(* IEC 61131-3 sources: daoli-st-library/DL_Motion (part 20) *)

(* ---- FB_DL_UnwinderDiameterCalc.st ---- *)
(*==============================================================================
 * 组件名称 (Component)  : FB_DL_UnwinderDiameterCalc
 * 所属子库 (Sublibrary) : DL_Motion
 * 当前版本 (Version)    : 1.0.0
 * 兼容性 (Platform)     : CODESYS 3.5 / TwinCAT 3 / 汇川 InoProShop / Machine Expert
 *                         仅依赖纯 IEC 61131-3 标准元素，零厂商方言
 * 功能描述 (Function)   : 放卷卷径实时估算：fDia = sqrt(fDiaInit^2 - 4 x thick x
 *                         SigmaLen / pi)，开方委托 FC_DL_NthRoot(2)；按外部累计
 *                         放膜长度增量递推；低于最小卷径 → bSpoolEnd 预警。
 *                         被开方数 < 0（数据矛盾）→ 冻结并报错，不塞伪值。
 * 溯源 (Origin)         : 道莅 clean-room 防御性实现
 * 本文件内含 (Contains) : TYPE E_DL_UnwdErr / FUNCTION_BLOCK FB_DL_UnwinderDiameterCalc
 * 依赖 (Depends)        : DL_MathData/FC_DL_NthRoot
 * 红线自检 (Redline)    : 无外部全局变量、无硬件地址直引 ｜ 全变量中英双语同行注释
 *                         防除零 + 量程钳位 + 非有限值防御 ｜ 枚举成员全部显式赋值
 *                         开方委托不重实现 ｜ 浮点容差比较 ｜ 输出冻结语义显式
 * 错误码表 (Codes)      : 16#0004_0318 就绪
 *                         16#0004_0319 信息级 膜厚非法(已钳制下限)
 *                         16#0004_031A 故障级 长度增量非法(拒绝递推)
 *                         16#0004_031B 故障级 数据矛盾(根号内负值或非有限，冻结输出)
 *                         16#0004_031C 信息级 接近空卷预警
 * 修订历史 (Revision)   : 2026-11-17  v1.0.0  首版入库 · R27 · 阶段三批 3
 * 验收向量 (Acceptance) : 初始卷径 500 mm，膜厚 50 um，累计放膜 1000 m
 *                         → 卷径 = sqrt(500^2 - 4*0.05*1000/3.14159...) ≈ 499.94 mm
 *============================================================================*)

(*-----------------------------------------------------------------------------
 * 枚举: E_DL_UnwdErr（归属 DL_Motion，与 FB_DL_UnwinderDiameterCalc 同文件）
 *----------------------------------------------------------------------------*)
TYPE E_DL_UnwdErr :
(
    eReady      := 16#0004_0318,   // 就绪 / Ready
    eThickClamp := 16#0004_0319,   // 信息级：膜厚非法已钳制下限 / Info: film thickness clamped
    eLenIncrBad := 16#0004_031A,   // 故障级：长度增量非法（放卷长度不允许回退）/ Fault: illegal length increment
    eDataContrad:= 16#0004_031B,   // 故障级：数据矛盾（根号内负值或非有限，冻结）/ Fault: data contradiction, output frozen
    eSpoolEnd   := 16#0004_031C    // 信息级：接近空卷预警 / Info: spool-end warning
);
END_TYPE

(*==============================================================================
 * 功能块: FB_DL_UnwinderDiameterCalc
 * 调用约定: 每个扫描周期无条件调用一次；fWebLen_m 必须为单调不减的累计放膜长度。
 *============================================================================*)
FUNCTION_BLOCK FB_DL_UnwinderDiameterCalc
VAR_INPUT
    fFilmThick_um : REAL;              // 膜厚 [微米]，有效域 5~500 / Film thickness [um]
    fDiaInit_mm   : REAL;              // 初始卷径 [毫米]，有效域 50~1200 / Initial roll diameter [mm]
    fWebLen_m     : REAL;              // 累计放膜长度 [米]（外部积分输入，单调不减）/ Accumulated web length [m]
    fDiaMin_mm    : REAL;              // 最小卷径 [毫米]（空卷预警门限）/ Minimum roll diameter [mm]
    bReset        : BOOL;              // 换卷复位（重新以初始卷径起算）/ Roll-change reset
END_VAR
VAR_OUTPUT
    fDiaNow_mm    : REAL;              // 当前卷径 [毫米] / Current roll diameter [mm]
    bSpoolEnd     : BOOL;              // 接近空卷预警 / Spool-end warning
    eErr          : E_DL_UnwdErr;      // 错误码 / Error code
END_VAR
VAR
    fLenPrev      : REAL;              // 上拍累计长度快照 [米]（增量基准）/ Previous length snapshot [m]
    fLenUse       : REAL;              // 生效累计长度（增量非法时冻结）[米] / Effective accumulated length [m]
    fThickUse_mm  : REAL;              // 生效膜厚（换算毫米，钳位后）[毫米] / Effective thickness in mm [mm]
    fDiaInitUse   : REAL;              // 生效初始卷径（NaN 兜底）[毫米] / Effective initial diameter [mm]
    fLenIncr      : REAL;              // 本拍长度增量 [米] / Length increment this scan [m]
    fRadicand     : LREAL;             // 被开方数 [平方毫米] / Radicand [mm2]
    fRootVal      : LREAL;             // 委托开方输出 [毫米] / Delegate root output [mm]
    bRootOk       : BOOL;              // 委托开方有效标志 / Delegate root validity flag
    bFrozen       : BOOL;              // 输出冻结标志（数据矛盾置位）/ Output frozen flag
    bInit         : BOOL;              // 首扫初始化标志 / First-scan init flag
END_VAR
VAR CONSTANT
    DL_UNWD_THICK_MIN : REAL := 5.0;      // 膜厚下限 [微米] / Thickness lower bound [um]
    DL_UNWD_THICK_MAX : REAL := 500.0;    // 膜厚上限 [微米] / Thickness upper bound [um]
    DL_UNWD_DIA_MIN   : REAL := 50.0;     // 初始卷径下限 [毫米] / Initial diameter lower bound [mm]
    DL_UNWD_DIA_MAX   : REAL := 1200.0;   // 初始卷径上限 [毫米] / Initial diameter upper bound [mm]
    DL_UNWD_UM2MM     : REAL := 0.001;    // 微米换毫米系数 [毫米每微米] / um-to-mm factor [mm per um]
    DL_UNWD_M2MM      : REAL := 1000.0;   // 米换毫米系数 [毫米每米] / m-to-mm factor [mm per m]
    DL_UNWD_FOUR      : REAL := 4.0;      // 面积递推系数 4（4 x thick x len / pi）/ Area recursion factor
    DL_UNWD_PI        : REAL := 3.14159265358979;   // 圆周率 [无量纲] / Pi [dimensionless]
    DL_UNWD_TOL       : REAL := 1.0E-6;   // 浮点比较容差 / Float comparison tolerance
    DL_UNWD_INF_MAX   : REAL := 1.0E30;   // 非有限值判定幅值上限 / Magnitude bound for finite-value check
    DL_UNWD_ZERO      : REAL := 0.0;      // 零值常量，避免裸字面量 / Zero constant
END_VAR

(*------------------------------------------------------------------------------
 * 段 1｜换卷复位：清快照与冻结标志，卷径回初始值
 *----------------------------------------------------------------------------*)
IF bReset THEN
    fLenPrev := fWebLen_m;                         // 快照重置为当前累计长度 / snapshot reset
    fLenUse := fWebLen_m;                          // 累计长度重置 / length reset
    fDiaNow_mm := fDiaInit_mm;                     // 卷径回初始值 / diameter back to initial
    bFrozen := FALSE;                              // 冻结解除 / freeze released
    bSpoolEnd := FALSE;                            // 预警解除 / warning released
    bInit := TRUE;                                 // 视为首扫完成（跳过旧快照）/ treated as initialized
    eErr := E_DL_UnwdErr.eReady;                   // 回就绪码 / back to ready
    RETURN;
END_IF

(*------------------------------------------------------------------------------
 * 段 2｜首扫初始化：建立长度快照基准
 *----------------------------------------------------------------------------*)
IF NOT bInit THEN
    fLenPrev := fWebLen_m;                         // 首扫快照 / first-scan snapshot
    fLenUse := fWebLen_m;                          // 累计长度基准 / length baseline
    bInit := TRUE;                                 // 首扫完成 / first scan done
END_IF

(*------------------------------------------------------------------------------
 * 段 3｜非有限值闸：任一输入 NaN/溢出 → 冻结输出并报数据矛盾（不塞伪值）
 *----------------------------------------------------------------------------*)
IF (fFilmThick_um <> fFilmThick_um) OR (ABS(fFilmThick_um) > DL_UNWD_INF_MAX)
   OR (fDiaInit_mm <> fDiaInit_mm) OR (ABS(fDiaInit_mm) > DL_UNWD_INF_MAX)
   OR (fWebLen_m <> fWebLen_m) OR (ABS(fWebLen_m) > DL_UNWD_INF_MAX)
   OR (fDiaMin_mm <> fDiaMin_mm) OR (ABS(fDiaMin_mm) > DL_UNWD_INF_MAX) THEN
    bFrozen := TRUE;                               // 输出冻结 / output frozen
    eErr := E_DL_UnwdErr.eDataContrad;             // 故障级：数据矛盾（非有限并入）/ fault: data contradiction
    bSpoolEnd := TRUE;                             // 数据矛盾按安全侧预警 / safe-side warning
    RETURN;
END_IF

(*------------------------------------------------------------------------------
 * 段 4｜膜厚钳位（信息级）与初始卷径兜底
 *----------------------------------------------------------------------------*)
eErr := E_DL_UnwdErr.eReady;                       // 预置就绪 / preset ready
fThickUse_mm := fFilmThick_um * DL_UNWD_UM2MM;     // 膜厚换算毫米 [毫米] / thickness to mm
IF fFilmThick_um < DL_UNWD_THICK_MIN THEN
    fThickUse_mm := DL_UNWD_THICK_MIN * DL_UNWD_UM2MM;   // 膜厚下限钳制 / thickness floored
    eErr := E_DL_UnwdErr.eThickClamp;              // 信息级：膜厚非法已钳制 / info: thickness clamped
ELSIF fFilmThick_um > DL_UNWD_THICK_MAX THEN
    fThickUse_mm := DL_UNWD_THICK_MAX * DL_UNWD_UM2MM;   // 膜厚上限钳制 / thickness capped
    eErr := E_DL_UnwdErr.eThickClamp;              // 信息级：膜厚非法已钳制 / info: thickness clamped
END_IF
fDiaInitUse := fDiaInit_mm;                        // 初始卷径工作副本 / initial diameter working copy
IF (fDiaInitUse < DL_UNWD_DIA_MIN) OR (fDiaInitUse > DL_UNWD_DIA_MAX) THEN
    fDiaInitUse := DL_UNWD_DIA_MIN;                // 初始卷径出域按下限兜底（配置防御）/ initial diameter falls back
END_IF

(*------------------------------------------------------------------------------
 * 段 5｜长度增量合法性闸：放卷长度单调不减（容差内视为零增量）
 *----------------------------------------------------------------------------*)
fLenIncr := fWebLen_m - fLenPrev;                  // 本拍增量 [米] / increment this scan [m]
IF fLenIncr < -DL_UNWD_TOL THEN
    bFrozen := TRUE;                               // 增量为负：拒绝递推，冻结输出 / negative increment: reject, freeze
    eErr := E_DL_UnwdErr.eLenIncrBad;              // 故障级：长度增量非法 / fault: illegal increment
    fLenUse := fLenPrev;                           // 冻结到上拍快照 / frozen at previous snapshot
    RETURN;
END_IF
IF fLenIncr < DL_UNWD_ZERO THEN
    fLenIncr := DL_UNWD_ZERO;                      // 容差内微负增量钳零 / tiny negative clamped to zero
END_IF
fLenUse := fLenPrev + fLenIncr;                    // 生效累计长度 [米] / effective length [m]
fLenPrev := fWebLen_m;                             // 快照推进 / snapshot advanced

(*------------------------------------------------------------------------------
 * 段 6｜卷径递推：被开方数 = 初始卷径^2 - 4 x 膜厚 x 累计长度 / pi
 *       被开方数 < 0（数据矛盾：放膜量超过卷料面积）→ 冻结并报故障级
 *----------------------------------------------------------------------------*)
fRadicand := REAL_TO_LREAL(fDiaInitUse * fDiaInitUse)
           - REAL_TO_LREAL(DL_UNWD_FOUR * fThickUse_mm * fLenUse * DL_UNWD_M2MM) / REAL_TO_LREAL(DL_UNWD_PI);   // 被开方数 [平方毫米]（米换毫米链）/ radicand [mm2]
IF (fRadicand <> fRadicand) OR (ABS(fRadicand) > REAL_TO_LREAL(DL_UNWD_INF_MAX)) THEN
    bFrozen := TRUE;                               // 非有限中间量：冻结 / non-finite intermediate: freeze
    eErr := E_DL_UnwdErr.eDataContrad;             // 故障级：数据矛盾 / fault: data contradiction
    bSpoolEnd := TRUE;                             // 安全侧预警 / safe-side warning
    RETURN;
END_IF
IF fRadicand < LREAL#0.0 THEN
    bFrozen := TRUE;                               // 根号内负值：数据矛盾冻结 / negative radicand: freeze
    eErr := E_DL_UnwdErr.eDataContrad;             // 故障级：根号内负值 / fault: negative radicand
    bSpoolEnd := TRUE;                             // 安全侧预警 / safe-side warning
    RETURN;
END_IF

(*------------------------------------------------------------------------------
 * 段 7｜委托开方（FC_DL_NthRoot(2)）与空卷预警
 *----------------------------------------------------------------------------*)
fRootVal := FC_DL_NthRoot(fValue := fRadicand, nRoot := 2, bValid => bRootOk);   // 开方委托 [毫米] / root via delegate [mm]
IF (NOT bRootOk) OR (fRootVal <> fRootVal) OR (ABS(fRootVal) > REAL_TO_LREAL(DL_UNWD_INF_MAX)) THEN
    bFrozen := TRUE;                               // 委托失败：冻结 / delegate failure: freeze
    eErr := E_DL_UnwdErr.eDataContrad;             // 故障级：数据矛盾（委托失败并入，输出同为冻结）/ fault: contradiction
    RETURN;
END_IF
fDiaNow_mm := LREAL_TO_REAL(fRootVal);             // 当前卷径输出 [毫米] / current diameter output [mm]
IF fDiaNow_mm < DL_UNWD_ZERO THEN
    fDiaNow_mm := DL_UNWD_ZERO;                    // 下限防护 / floor guard
END_IF
bSpoolEnd := fDiaNow_mm <= fDiaMin_mm + DL_UNWD_TOL;   // 空卷预警判据（容差比较）/ spool-end predicate
IF bSpoolEnd THEN
    eErr := E_DL_UnwdErr.eSpoolEnd;                // 信息级：接近空卷 / info: spool-end warning
END_IF
END_FUNCTION_BLOCK

(* ---- FB_DL_VelFfGainIdent.st ---- *)
(*==============================================================================
 * 组件名称 (Component)  : FB_DL_VelFfGainIdent
 * 所属子库 (Sublibrary) : DL_Motion
 * 当前版本 (Version)    : 1.0.0
 * 兼容性 (Platform)     : CODESYS 3.5+ / TwinCAT 3 / 汇川 InoProShop / 施耐德 Machine Expert
 *                         仅依赖 Standard.library（TON / R_TRIG），零厂商私有库，
 *                         零轴状态枚举引用（R277）
 * 功能描述 (Function)   : 速度前馈增益辨识。恒速段窗口（bConstVel 电平：上层
 *                         速度指令平坦段）内对 (vFb, vCmd) 做 最小二乘 过原点
 *                         拟合 K = Σ(vFb·vCmd) / Σ(vFb²)（前馈模型 vCmd ≈ K·vFb
 *                         的残差最优解），同步累计残差标准差与样本数；样本充分
 *                         且拟合优度高（残差/信号比小）→ bIdentDone 单拍输出
 *                         fKvf。与 AxisFrictionFf 分工：本件辨识增益不注入
 *                         前馈（R312 模型不内嵌注入语义）。
 * 来源标签 (Origin)     : 自研线（IEC 61131-3 标准语义的道莅防御性实现，clean-room）
 * 分工声明 (Pairing)    : VelFfGainIdent（辨识，本件）↔ AxisFrictionFf（前馈注入，
 *                         既有件）：本件只产出辨识增益与置信指标，不写前馈通道、
 *                         不驱动轴（R298 属主边界）；辨识结果由调用方决定是否
 *                         下装（R312 口径）。
 * 边界语义 (Boundary)   : ① 过原点拟合分母闸：Σ(vFb²) <= eps（恒速段实际零速
 *                         或样本未采）→ 拟合不执行，K 保持上值；
 *                         ② 速度非有限拒收（NaN 自反 + Inf 差判）；
 *                         ③ 置信闸：残差均方根/均值 |vCmd| > fConfRatio
 *                         → 拟合质量不足，bIdentDone 不置位（辨识不可信
 *                         必须可观测，R28 口径）；
 *                         ④ 组态闸：最小样本/置信比/增益钳位域 → 故障。
 * 输出语义 (Fallback)   : 【R191】bConstVel = FALSE → 停止采样，fKvf 保持
 *                         末次辨识值（增益是资产，不随窗口停而清零）；
 *                         eFault 相 → 冻结 + bError = TRUE。
 * 码位     (Codes)      : 按 R297 范式零 16# 码位硬编码；错误出口 BOOL+ENUM(eCause)，
 *                         码位待主控收口统一派号。
 * 红线自检 (Redline)    : 7 项红线已自检：R1 零全局 ✓｜R2 零物理地址 ✓｜R3 纯 IEC ✓
 *                         R4 除零（Σv² eps 闸）/NaN 拒收/组态闸 ✓
 *                         R5 双语同行注释 ✓｜R6 CASE 带 ELSE 兜底迁 eFault ✓
 *                         R7 TON/R_TRIG 段 0 无条件刷新 ✓
 * 验收向量 (Acceptance) : V1 恒速段 vCmd=vFb=200 → K=1.0（容差 1E-6）；
 *                         V2 vFb 恒为 vCmd 的 0.8 倍 → K=1.25；
 *                         V3 零速恒速段（vFb≈0）→ 分母闸生效，K 保持上值；
 *                         V4 残差比超阈 → bIdentDone 不置位。
 * 修订历史 (Revision)   : 2026-11-20  v1.0.0  R49 首版（批 4 · 序号 17）
 *==============================================================================*)
TYPE E_DL_VfiState :
(
    eIdle  := 0,                             (* 待使能 / Idle *)
    eLearn := 10,                            (* 恒速段采样与拟合 / Learning *)
    eFault := 90                             (* 故障锁存相 / Fault latched phase *)
);
END_TYPE

TYPE E_DL_VfiCause :
(
    eNone       := 0,                        (* 无故障成因 / No cause *)
    eCfgIllegal := 1,                        (* 组态非法：样本/置信比越域 / Illegal config *)
    ePhaseBad   := 2                         (* 非法相位兜底 / Illegal phase fallback *)
);
END_TYPE

FUNCTION_BLOCK FB_DL_VelFfGainIdent
VAR_INPUT
    fVelCmd    : LREAL := 0.0;               (* 速度指令反馈快照 [mm/s] / Velocity command snapshot *)
    fVelFb     : LREAL := 0.0;               (* 实际速度反馈快照 [mm/s] / Velocity feedback snapshot *)
    bConstVel  : BOOL := FALSE;              (* 恒速段电平（上层速度平坦段判据直连）[-] / Constant-velocity window level *)
    nMinSample : INT := 64;                  (* 最小辨识样本数，域 8..100000 [点] / Min identification samples *)
    fConfRatio : LREAL := 0.1;               (* 置信比门限（残差 RMS / 均值|vCmd|），域 (0,1) [-] / Confidence ratio gate *)
    bEnable    : BOOL := TRUE;               (* 辨识使能 [-] / Enable *)
    bReset     : BOOL := FALSE;              (* 复位命令，上升沿清累计与锁存（fKvf 保留）[-] / Reset command *)
END_VAR
VAR_OUTPUT
    fKvf       : LREAL;                      (* 辨识速度前馈增益（末次有效值保持）[-] / Identified velocity ff gain *)
    nSampleCnt : INT;                        (* 本轮累计样本数 [点] / Sample count this round *)
    fResidRms  : LREAL;                      (* 跟随残差均方根（拟合质量）[mm/s] / Residual RMS *)
    bIdentDone : BOOL;                       (* 本轮辨识完成单拍位（质量闸通过才置位）[-] / Round-done single-scan pulse *)
    bIdentFail : BOOL;                       (* 本轮辨识质量不足锁存位（复位沿清）[-] / Round-quality-fail latch *)
    eState     : E_DL_VfiState;              (* 状态出口 / State outlet *)
    eCause     : E_DL_VfiCause;              (* 故障成因出口（R190 归因唯一） / Fault cause outlet *)
    bError     : BOOL;                       (* 故障锁存标志 [-] / Fault latch flag *)
END_VAR
VAR
    _eState  : E_DL_VfiState := E_DL_VfiState.eIdle;      (* 内部相位（CASE 唯一写入目标） / Internal phase *)
    _eCause  : E_DL_VfiCause := E_DL_VfiCause.eNone;      (* 故障成因锁存量 / Latched cause *)
    rtReset  : R_TRIG;                       (* 复位沿实例，段 0 无条件调用 / Reset edge instance *)
    _nCnt    : INT;                          (* 样本计数锁存 [点] / Sample count latch *)
    _nMin    : INT;                          (* 钳位后生效最小样本数 [点] / Clamped min samples *)
    _fSfb2   : LREAL;                        (* Σ vFb² 累计 [mm²/s²] / Sum of vFb squared *)
    _fSfbc   : LREAL;                        (* Σ vFb·vCmd 累计 [mm²/s²] / Sum of vFb·vCmd *)
    _fSres2  : LREAL;                        (* Σ 残差² 累计（按上轮 K 算的即时残差）[mm²/s²] / Sum of squared residual *)
    _fSumAbs : LREAL;                        (* Σ |vCmd| 累计（置信比分母）[mm/s] / Sum of |vCmd| *)
    _fK      : LREAL := 1.0;                 (* 拟合增益锁存（缺省 1.0 = 无前馈修正语义）[-] / Fitted gain latch *)
    _bFault  : BOOL;                         (* 故障锁存位 / Latched fault bit *)
    _bCfgBad : BOOL;                         (* 组态非法当拍量 / Illegal config this scan *)
END_VAR
VAR CONSTANT
    DL_VFI_EPS : LREAL := 1.0E-9;            (* 拟合分母判零容差 [mm²/s²] / Fit denominator epsilon *)
    DL_VFI_NMAX: INT   := 100000;            (* 样本上限（防 INT 溢出）[点] / Sample upper limit *)
    DL_VFI_KMAX: LREAL := 10.0;              (* 增益钳位上限（异常拟合兜底，R151 口径）[-] / Gain clamp limit *)
    DL_VFI_KMIN: LREAL := 0.1;               (* 增益钳位下限 [-] / Gain clamp lower limit *)
END_VAR

(* —— 段 0：当拍判据派生 + 实例无条件刷新（R228A） —— *)
_bCfgBad := (nMinSample < 8) OR (nMinSample > DL_VFI_NMAX) OR (fConfRatio <= 0.0) OR (fConfRatio >= 1.0);   (* 组态闸（R151 全引脚） / Config gate *)
rtReset(CLK := bReset);                      (* 复位沿每拍必调 / Reset edge every scan *)
_nMin := nMinSample;                         (* 生效最小样本初值 / Min init *)
IF _nMin < 8 THEN
    _nMin := 8;                              (* 下限钳位 / Lower clamp *)
END_IF
IF _nMin > DL_VFI_NMAX THEN
    _nMin := DL_VFI_NMAX;                    (* 上限钳位（R308） / Upper clamp *)
END_IF

(* —— 段 1：单拍量预清零（R107） —— *)
bIdentDone := FALSE;                         (* 完成单拍位预清，唯一分支置位 / Done pulse preset *)

(* —— 段 2：复位沿处理（作用域：清故障 + 清全部累计量 + 清样本数 + 清质量锁存；fKvf 保留，R283 逐项声明） —— *)
IF rtReset.Q THEN
    _bFault := FALSE;                        (* 清故障锁存 / Clear fault *)
    _eCause := E_DL_VfiCause.eNone;          (* 清成因 / Clear cause *)
    _nCnt := 0;                              (* 清样本数 / Clear count *)
    _fSfb2 := 0.0;                           (* 清 ΣvFb² / Clear sum *)
    _fSfbc := 0.0;                           (* 清 ΣvFb·vCmd / Clear sum *)
    _fSres2 := 0.0;                          (* 清 Σ残差² / Clear sum *)
    _fSumAbs := 0.0;                         (* 清 Σ|vCmd| / Clear sum *)
    fResidRms := 0.0;                        (* 清 RMS 出口 / Clear outlet *)
    bIdentFail := FALSE;                     (* 清质量不足锁存 / Clear fail latch *)
    nSampleCnt := 0;                         (* 清样本出口 / Clear count outlet *)
    _eState := E_DL_VfiState.eIdle;          (* 迁待机相 / Back to idle *)
END_IF

(* —— 段 3：组态闸故障锁存（R45 配对；锁存至复位沿，R189） —— *)
IF _bCfgBad AND NOT _bFault THEN
    _bFault := TRUE;                         (* 锁存故障位 / Latch fault *)
    _eCause := E_DL_VfiCause.eCfgIllegal;    (* 成因：组态非法 / Cause: illegal config *)
    _eState := E_DL_VfiState.eFault;         (* 同步迁故障相 / Migrate to fault *)
END_IF

(* —— 段 4：CASE 主状态机（ELSE 兜底迁 eFault，红线 6） —— *)
CASE _eState OF
    E_DL_VfiState.eIdle:                     (* 待机相 / Idle *)
        IF bEnable AND NOT _bFault THEN
            _eState := E_DL_VfiState.eLearn; (* 进入学习 / Enter learn *)
        END_IF
    E_DL_VfiState.eLearn:                    (* 学习相：恒速段采样 + 过原点 LS 拟合 / Learn *)
        IF NOT bEnable THEN
            _eState := E_DL_VfiState.eIdle;  (* 失能回待机（fKvf 保持） / Back to idle *)
        ELSIF bConstVel THEN                 (* 仅恒速段采样（判据串相位因子，R281） / Sample only in const-vel *)
            IF (fVelFb = fVelFb) AND (fVelCmd = fVelCmd)
               AND ((fVelFb - fVelFb) = (fVelFb - fVelFb)) AND ((fVelCmd - fVelCmd) = (fVelCmd - fVelCmd)) THEN
                _fSfb2 := _fSfb2 + fVelFb * fVelFb;       (* ΣvFb² 累计 / Accumulate *)
                _fSfbc := _fSfbc + fVelFb * fVelCmd;      (* ΣvFb·vCmd 累计 / Accumulate *)
                _fSres2 := _fSres2 + (fVelCmd - _fK * fVelFb) * (fVelCmd - _fK * fVelFb);   (* 即时残差² 累计（按当前 K） / Instant residual² *)
                _fSumAbs := _fSumAbs + ABS(fVelCmd);      (* Σ|vCmd| 累计 / Accumulate *)
                IF _nCnt < DL_VFI_NMAX THEN
                    _nCnt := _nCnt + 1;      (* 样本计数（INT 溢出防护） / Count advance *)
                END_IF
            END_IF
            IF _fSfb2 > DL_VFI_EPS THEN      (* 分母闸：恒速段非零速才拟合（边界①） / Denominator gate *)
                _fK := _fSfbc / _fSfb2;      (* 过原点最小二乘 K = Σ(vFb·vCmd)/Σ(vFb²)（分母已过 eps 闸，无除零） / Origin-LS fit, denominator gated *)
                IF _fK > DL_VFI_KMAX THEN
                    _fK := DL_VFI_KMAX;      (* 增益上限钳位（异常拟合兜底） / Gain upper clamp *)
                ELSIF _fK < DL_VFI_KMIN THEN
                    _fK := DL_VFI_KMIN;      (* 增益下限钳位（IF 链带 ELSE 兜底，R285） / Gain lower clamp *)
                END_IF
            END_IF
            IF (_nCnt >= _nMin) AND (_fSfb2 > DL_VFI_EPS) AND (_nCnt >= 1) THEN
                fResidRms := SQRT(_fSres2 / INT_TO_LREAL(_nCnt));   (* RMS 出口（除子恒 >= 1，无除零） / RMS outlet *)
                IF ABS(fVelCmd) > DL_VFI_EPS OR _fSumAbs > DL_VFI_EPS THEN
                    IF (_fSumAbs / INT_TO_LREAL(_nCnt)) > DL_VFI_EPS AND (fResidRms / (_fSumAbs / INT_TO_LREAL(_nCnt))) <= fConfRatio THEN
                        fKvf := _fK;         (* 质量闸通过：增益下装出口 / Quality passed: gain outlet *)
                        bIdentDone := TRUE;  (* 完成单拍脉冲 / Done pulse *)
                        bIdentFail := FALSE; (* 清质量不足锁存 / Clear fail latch *)
                        _eState := E_DL_VfiState.eIdle;   (* 收口回待机（下轮重新累计） / Back to idle *)
                    ELSIF (_fSumAbs / INT_TO_LREAL(_nCnt)) > DL_VFI_EPS THEN
                        bIdentFail := TRUE;  (* 质量不足锁存至复位沿（R28 可观测口径） / Quality fail latch *)
                        _eState := E_DL_VfiState.eIdle;   (* 收口回待机 / Back to idle *)
                    END_IF
                END_IF
            END_IF
            nSampleCnt := _nCnt;             (* 样本数出口镜像 / Count mirror *)
        END_IF
    E_DL_VfiState.eFault:                    (* 故障相：冻结保持，仅复位沿出 / Fault *)
        ;                                    (* 锁存回放（R28） / Replay from latch *)
    ELSE                                     (* 非法相位兜底迁安全态 / Illegal phase fallback *)
        _eState := E_DL_VfiState.eFault;     (* 迁故障相 / To fault *)
        _bFault := TRUE;                     (* 同步锁存 / Latch *)
        _eCause := E_DL_VfiCause.ePhaseBad;  (* 成因：非法相位 / Cause: illegal phase *)
END_CASE

(* —— 段 5：出口映射（bError/eState 同源，R191） —— *)
bError := _bFault;                           (* 故障标志镜像 / Fault flag mirror *)
eState := _eState;                           (* 状态出口 / State outlet *)
eCause := _eCause;                           (* 成因出口 / Cause outlet *)
END_FUNCTION_BLOCK

(* ---- FB_DL_WaferCountAxis.st ---- *)
//==============================================================================
// 功能块：FB_DL_WaferCountAxis ｜ 中文名称：晶圆计数轴（编码器分频 + 片位同步）
// 所属子库：DL_Motion ｜ 版本：v1.0.0 ｜ 兼容：CODESYS V3.5+ / TwinCAT 3 / 汇川 InoProShop
// 功能描述：编码器脉冲分频晶圆计数——按脉冲/片分频比累计计片，片位同步
//           单拍脉冲输出（EAP 对账用），滑动窗估算节拍率 [片/min]。
// 开源溯源 (Origin)：道莅原创实现（参考半导体 EAP 对账与计数轴工程惯例 分类与参数域）
// 单位表：脉冲[—] / 分频比[脉冲/片] / 计数[片] / 节拍率[片/min] / 窗[ms]
// 错误码表：16#0004_01DF 信息级（计数饱和 4294967295，不回绕，不置
//           bError）/ 16#0004_01E0 预留禁用（不得挪用）/ 16#0004_02F9
//           故障级（分频比为 0，除零前置闸，置 bError）/ 16#0004_02FA
//           预留禁用（不得挪用）/ 16#0004_02FB 故障级兜底（置 bError）
// 状态机：N/A（分频计数 + 窗口估算为电平逻辑，无相位状态机）
// 边界行为：① uPulsesPerWafer = 0 → 故障 02F9（除零前置闸，计数冻结）；
//           ② 计数饱和 4294967295 + 信息 01DF，不回绕；③ bResetCount
//           优先级最高（同拍清分频累加器、窗计数与总计数）；④ 节拍率窗
//           tRateWindow <= 0 → 斜率走窗口为 0 的构造路径保护（估算率
//           冻结 0，不除零）；⑤ R_TRIG 首部无条件刷新（R40）。
// 依赖纪律：Motion 不得引用任何其他 DL_ 子库（R22 纪律延续）——本件仅用
//           Standard.library（TON/R_TRIG），未使用同库 I_DL_MotionAxis
//           （纯脉冲计数无需轴接口，头注释声明此设计取舍）。
// 修订历史：v1.0.0 2026-11-17 首版（R23 派单 · ROADMAP 半导体 P1 §369）
//==============================================================================

FUNCTION_BLOCK FB_DL_WaferCountAxis
VAR_INPUT
    bEncPulse       : BOOL;                 // 编码器脉冲输入 [—] / Encoder pulse input
    uPulsesPerWafer : UINT := 100;          // 分频比 [脉冲/片]，须 > 0 / Divider ratio [pulses per wafer], must be > 0
    bCountEnable    : BOOL;                 // 计数使能 [—] / Count enable
    bResetCount     : BOOL;                 // 计数复位 [—]，优先级最高 / Count reset, highest priority
END_VAR
VAR_OUTPUT
    uWaferCount     : UDINT;                // 晶圆计数 [片]，饱和 4294967295 不回绕 / Wafer count [pieces], saturated without wrap
    bWaferIndexPulse: BOOL;                 // 片位同步单拍脉冲 [—] / Wafer-index one-scan pulse
    fEstRate        : LREAL;                // 估算节拍率 [片/min] / Estimated rate [pieces/min]
    eErr            : UDINT;                // 错误码，0 = 无错 / Error code, 0 = no error
    bError          : BOOL;                 // 故障级标志，仅故障级错误置位 / Fault-class flag, set only on fault-level codes
    bValid          : BOOL;                 // 输出可用标志 / Outputs usable flag
END_VAR
VAR
    rtEnc           : R_TRIG;               // 编码器脉冲上升沿，段 6 无条件刷新 / Encoder pulse rising edge
    fbRateWin       : TON;                  // 节拍率估算窗，段 6 无条件刷新 [ms] / Rate estimation window
    _uPulseAcc      : UINT;                 // 分频脉冲累加器 [脉冲] / Divider pulse accumulator [pulses]
    _uWinCount      : UINT;                 // 窗内计片数 [片] / Wafer count within the window [pieces]
    _fWinMinutes    : LREAL;                // 估算窗时长 [min] / Window duration [min]
    _bInit          : BOOL := FALSE;        // 首扫标志，初值 FALSE 取非判定 / First-scan flag, tested negated
    _bDivZero       : BOOL;                 // 分频比为 0 锁存 / Zero-divider latch
    _bSaturated     : BOOL;                 // 计数饱和当拍标志 / Saturation flag of this scan
    _bIdxPulse      : BOOL;                 // 片位脉冲单拍标志 / One-scan index pulse flag
END_VAR
VAR CONSTANT
    DL_WC_CNT_MAX   : UDINT := 4294967295;  // 计数饱和上限 [片] / Counter saturation ceiling [pieces]
    DL_WC_RATE_WIN  : TIME  := T#10S;       // 节拍率估算窗 [ms] / Rate estimation window [ms]
    DL_WC_MS_PER_MIN: LREAL := 60000.0;     // 毫秒 → 分钟换算系数 [ms/min] / Millisecond-to-minute factor [ms/min]
    DL_WC_INF       : LREAL := 1.7976931348623157E308; // LREAL 幅值上限 / LREAL magnitude ceiling
END_VAR

(*------------------------------------------------------------------------------
 * 段 1｜每拍预置：输出先算后出，单拍标志预清零（R25 第一律：只置必销）
 *      Outputs computed per scan, one-shot flags pre-cleared
 *-----------------------------------------------------------------------------*)
bWaferIndexPulse := FALSE;                  // 片位脉冲预清零 / Index pulse pre-cleared
fEstRate         := 0.0;                    // 节拍率预置零 / Rate preset zero
eErr             := 16#0000_0000;           // 错误码每拍重算 / Error code recomputed
bError           := FALSE;                  // 故障标志每拍重算 / Fault flag recomputed
bValid           := FALSE;                  // 可用标志每拍重算 / Usable flag recomputed
_bSaturated      := FALSE;                  // 饱和标志预清零 / Saturation flag pre-cleared
_bIdxPulse       := FALSE;                  // 片位暂存预清零 / Index staging pre-cleared

(*------------------------------------------------------------------------------
 * 段 2｜首扫初始化
 *      First-scan initialisation
 *-----------------------------------------------------------------------------*)
IF NOT _bInit THEN
    uWaferCount := 0;                       // 计数清零 / Counter cleared
    _uPulseAcc  := 0;                       // 分频累加器清零 / Accumulator cleared
    _uWinCount  := 0;                       // 窗计数清零 / Window counter cleared
    _bDivZero   := FALSE;                   // 除零锁存清零 / Zero-divider latch cleared
    _bInit      := TRUE;                    // 首扫只做一次 / The first scan runs once
END_IF

(*------------------------------------------------------------------------------
 * 段 3｜R_TRIG 与估算窗无条件刷新（R40：CASE 之外每拍必调）
 *      R_TRIG and the rate window refreshed unconditionally per R40
 *-----------------------------------------------------------------------------*)
rtEnc(CLK := bEncPulse);                    // 编码器脉冲上升沿 / Encoder pulse rising edge
fbRateWin(IN := bCountEnable AND (NOT _bDivZero), PT := DL_WC_RATE_WIN); // 节拍率估算窗 / Rate estimation window

(*------------------------------------------------------------------------------
 * 段 4｜复位优先级最高：清全部累计量
 *      Reset has the highest priority, clears every accumulator
 *-----------------------------------------------------------------------------*)
IF bResetCount THEN
    uWaferCount := 0;                       // 总计数清零 / Counter cleared
    _uPulseAcc  := 0;                       // 分频累加器清零 / Accumulator cleared
    _uWinCount  := 0;                       // 窗计数清零 / Window counter cleared
END_IF

(*------------------------------------------------------------------------------
 * 段 5｜分频计数：使能 + 沿有效时累加，达分频比进片（计数饱和不回绕）
 *      Divider counting with saturation guard
 *-----------------------------------------------------------------------------*)
IF bCountEnable AND (NOT _bDivZero) AND rtEnc.Q AND (NOT bResetCount) THEN
    IF _uPulseAcc + 1 >= uPulsesPerWafer THEN
        _uPulseAcc := 0;                    // 分频累加器归零 / Accumulator rolled over
        IF uWaferCount < DL_WC_CNT_MAX THEN
            uWaferCount := uWaferCount + 1; // 计片递增 / Wafer count increment
            _uWinCount  := _uWinCount + 1;  // 窗计数递增 / Window counter increment
            _bIdxPulse := TRUE;             // 片位脉冲单拍置位（段 1 预清，只置必销） / One-scan index pulse
        ELSE
            _bSaturated := TRUE;            // 计数饱和声明 / Saturation declared
        END_IF
    ELSE
        _uPulseAcc := _uPulseAcc + 1;       // 分频累加 / Accumulator increment
    END_IF
END_IF

(*------------------------------------------------------------------------------
 * 段 6｜节拍率估算：窗满按窗计片换算 [片/min]（窗 <= 0 走构造路径冻结）
 *      Rate estimation with the zero-window construction-path guard
 *-----------------------------------------------------------------------------*)
_fWinMinutes := TIME_TO_DINT(DL_WC_RATE_WIN) / DL_WC_MS_PER_MIN; // 窗时长 [min] / Window duration [min]
IF fbRateWin.Q AND (_fWinMinutes > 0.0) THEN
    fEstRate := UINT_TO_LREAL(_uWinCount) / _fWinMinutes; // 节拍率 [片/min]（标准类型转换，零方言） / Estimated rate [pieces/min], standard conversion
    _uWinCount := 0;                        // 窗计数清零重开 / Window counter cleared and restarted
END_IF

(*------------------------------------------------------------------------------
 * 段 7｜组态闸与码位出口
 *      Configuration gate and the code outlet
 *-----------------------------------------------------------------------------*)
IF uPulsesPerWafer = 0 THEN
    _bDivZero := TRUE;                      // 除零前置闸锁存（计数冻结） / Zero-divider latch, counting frozen
END_IF
bWaferIndexPulse := _bIdxPulse;             // 片位脉冲出口 / Index pulse outlet

IF _bDivZero THEN
    eErr   := 16#0004_02F9;                 // 故障级：分频比为 0 / Fault: zero divider ratio
    bError := TRUE;                         // 置故障标志（R45 配对） / Raise the fault flag
    bValid := FALSE;                        // 输出不可用 / Outputs unusable
ELSIF _bSaturated THEN
    eErr := 16#0004_01DF;                   // 信息级：计数饱和不回绕 / Info: counter saturated without wrap
    bValid := TRUE;                         // 输出可用 / Outputs usable
ELSE
    bValid := bCountEnable;                 // 使能且正常：输出可用 / Outputs usable when enabled
END_IF
END_FUNCTION_BLOCK

(* ---- FB_DL_WebGuideEpcSeq.st ---- *)
(*
  Component : FB_DL_WebGuideEpcSeq
  Category  : DL_Motion
  Function  : EPC 纠偏闭环状态机：找边扫描→跟踪（死区内不动）→丢边保持→换卷回中→故障锁存
  Complexity: C4
  开源溯源 : DLF 内部原创（R94 族模板派生）；参考语义来源见 SOURCE_HUNTING_MATRIX.md
  规则遵从 : R1-R16
  契约     : 输入 xStart 启动（上升沿启动，下降沿兼故障复位沿）、xStop 停止、xWebPresent 卷材存在、
             xSensorOk 传感器信号有效、xRollChange 换卷信号、rEdgeOffsetMm 边缘偏移（正=偏右） [mm]、
             rDeadbandMm 跟踪死区 [mm]、rFindBandMm 找边判定带宽 [mm]、rMaxOffsetMm 允许最大偏移 [mm]、
             rCorrRateMmS 跟踪纠偏速度 [mm/s]、rScanRateMmS 找边扫描速度 [mm/s]、
             rSearchTmoS 找边超时 [s]、rLostTmoS 丢边保持超时 [s]、rCenterTmoS 回中超时 [s]。
  输出     : rActCmdMmS 带符号执行速度指令（正=右移） [mm/s]、xMotionEnabled 执行使能、
             eState 当前相、xFault/nFaultCode 故障、nWarnCode 信息级码、xEdgeFound 已找到边。
  输出语义 : EDGE_LOST 相为「冻结保持末值」——执行速度指令保持进相前最后一拍的 rLastCmdMmS，
             设计理由：丢边瞬间若把指令清零会造成带材在纠偏辊上突然回弹（阶跃），
             故按冻结处理并在 nWarnCode 每拍报 9602，超时后转 FAULT 并强制撤销指令。
             xStop=TRUE 时不冻结，全部命令撤销并回 IDLE（撤销型停车）。
  复位沿   : 故障码锁存至 xStart 下降沿；复位后停在 IDLE，需重新给启动上升沿（不做自动再入）。
  码位     : 9601 找边超时（故障级）；9602 丢边保持中（信息级，不置 xFault）；
             9603 回中超时（故障级）；9604 参数或采样非法（故障级）；9605 卷材缺失（故障级）；
             9606 丢边保持超时（故障级，与 9601 分属不同成因，按 R190 归因唯一独立派码）。
*)
TYPE E_DL_WebGuideState :
(
    IDLE       := 0,    // 待机，执行使能撤销 EN: idle, the motion enable is withdrawn
    EDGE_SEARCH:= 10,   // 找边扫描相 EN: the edge search phase
    TRACKING   := 20,   // 跟踪相（死区内不动） EN: the tracking phase, no motion inside the dead band
    EDGE_LOST  := 30,   // 丢边保持相（指令冻结） EN: the edge lost phase with a frozen command
    CENTERING  := 40,   // 换卷回中相 EN: the centering phase after a roll change
    FAULT      := 90    // 故障相，指令强制撤销 EN: the fault phase, the command is forced off
);
END_TYPE

FUNCTION_BLOCK FB_DL_WebGuideEpcSeq
VAR_INPUT
    xStart        : BOOL;             // 启动（上升沿启动，下降沿复位故障） EN: start on the rising edge, reset the fault on the falling edge
    xStop         : BOOL;             // 停止（任意相生效，撤销指令） EN: stop, effective in every phase and withdrawing the command
    xWebPresent   : BOOL;             // 卷材存在（穿带完成） EN: the web is present after threading
    xSensorOk     : BOOL;             // 传感器信号有效 EDGE_LOST 判据 EN: the sensor signal is valid, the edge lost criterion
    xRollChange   : BOOL;             // 换卷信号（上升沿进回中相） EN: the roll change signal entering the centering phase
    rEdgeOffsetMm : REAL;             // 边缘偏移，正表示偏右 [mm] EN: the edge offset, positive means to the right
    rDeadbandMm   : REAL := 0.5;      // 跟踪死区 [mm] EN: the tracking dead band
    rFindBandMm   : REAL := 2.0;      // 找边判定带宽（进入该带即认为找到边） [mm] EN: the find band that declares an edge found
    rMaxOffsetMm  : REAL := 20.0;     // 允许最大偏移（越界视为异常） [mm] EN: the maximum allowed offset
    rCorrRateMmS  : REAL := 5.0;      // 跟踪纠偏速度幅值 [mm/s] EN: the tracking correction velocity magnitude
    rScanRateMmS  : REAL := 2.0;      // 找边扫描速度幅值 [mm/s] EN: the edge search velocity magnitude
    rSearchTmoS   : REAL := 30.0;     // 找边超时 [s] EN: the edge search timeout
    rLostTmoS     : REAL := 3.0;      // 丢边保持超时 [s] EN: the edge lost hold timeout
    rCenterTmoS   : REAL := 20.0;     // 回中超时 [s] EN: the centering timeout
END_VAR
VAR_OUTPUT
    rActCmdMmS    : REAL;             // 带符号执行速度指令，正表示右移 [mm/s] EN: the signed actuator velocity command, positive means right
    xMotionEnabled: BOOL;             // 执行使能 EN: the motion enable
    eState        : E_DL_WebGuideState;  // 当前相 EN: the current phase
    xFault        : BOOL;             // 故障标志（仅故障级码置位） EN: the fault flag, raised by fault class codes only
    nFaultCode    : INT;              // 故障码，锁存回放 EN: the fault code replayed from the latch
    nWarnCode     : INT;              // 信息级码（每拍重算） EN: the information class code recomputed every cycle
    xEdgeFound    : BOOL;             // 已找到边（跟踪相成立） EN: the edge has been found
END_VAR
VAR
    tonSearch  : TON;                 // 找边超时定时器 EN: the edge search timeout
    tonLost    : TON;                 // 丢边保持定时器 EN: the edge lost hold timer
    tonCenter  : TON;                 // 回中超时定时器 EN: the centering timeout
    fbStartRise: R_TRIG;              // xStart 上升沿（唯一启动沿） EN: the rising edge of xStart, the only start edge
    fbStartFall: F_TRIG;              // xStart 下降沿（复位沿） EN: the falling edge of xStart, the reset edge
    fbRollRise : R_TRIG;              // 换卷上升沿 EN: the rising edge of the roll change signal
    xFinAll    : BOOL;                // 全部浮点入参有限 EN: every floating input is finite
    xParamBad  : BOOL;                // 参数或采样非法 EN: a parameter or the sample is illegal
    xSensorUse : BOOL;                // 传感器可用（有效且偏移有限） EN: the sensor is usable
    rAbsOff    : REAL;                // 偏移绝对值 [mm] EN: the offset magnitude
    rCmd       : REAL;                // 本拍指令工作值 [mm/s] EN: the working command of this cycle
    rLastCmd   : REAL;                // 上拍指令快照（丢边冻结用） [mm/s] EN: the previous command snapshot used for the freeze
    nMsSearch  : UDINT := 30000;      // 找边超时毫秒数（缺省防零 PT） EN: the search timeout in milliseconds, the default avoids a zero preset
    nMsLost    : UDINT := 3000;       // 丢边超时毫秒数 EN: the lost timeout in milliseconds
    nMsCenter  : UDINT := 20000;      // 回中超时毫秒数 EN: the centering timeout in milliseconds
    nCodeLatch : INT;                 // 故障码锁存副本 EN: the latched copy of the fault code
END_VAR
VAR CONSTANT
    DL_WGE_Z       : REAL := 0.0;     // 浮点零常量 EN: the floating point zero constant
    DL_WGE_K1000   : REAL := 1000.0;  // 秒转毫秒系数 EN: the second to millisecond factor
    DL_WGE_W_LOST  : INT := 9602;     // 丢边保持中（信息级） EN: the edge is currently lost, information class
    DL_WGE_C_SEARCH: INT := 9601;     // 找边超时（故障级） EN: the edge search timed out
    DL_WGE_C_CENTER: INT := 9603;     // 回中超时（故障级） EN: the centering timed out
    DL_WGE_C_PARAM : INT := 9604;     // 参数或采样非法（故障级） EN: a parameter or the sample is illegal
    DL_WGE_C_WEB   : INT := 9605;     // 卷材缺失（故障级） EN: the web is missing
    DL_WGE_C_LOST  : INT := 9606;     // 丢边保持超时（故障级） EN: the edge lost hold timed out
END_VAR

// 段1｜参数与采样门禁（先判后用：换算在闸后，结果供段2 定时器 PT）
xFinAll := (rEdgeOffsetMm = rEdgeOffsetMm) AND ((rEdgeOffsetMm - rEdgeOffsetMm) = DL_WGE_Z)
        AND (rDeadbandMm = rDeadbandMm) AND ((rDeadbandMm - rDeadbandMm) = DL_WGE_Z)
        AND (rFindBandMm = rFindBandMm) AND ((rFindBandMm - rFindBandMm) = DL_WGE_Z)
        AND (rMaxOffsetMm = rMaxOffsetMm) AND ((rMaxOffsetMm - rMaxOffsetMm) = DL_WGE_Z)
        AND (rCorrRateMmS = rCorrRateMmS) AND ((rCorrRateMmS - rCorrRateMmS) = DL_WGE_Z)
        AND (rScanRateMmS = rScanRateMmS) AND ((rScanRateMmS - rScanRateMmS) = DL_WGE_Z)
        AND (rSearchTmoS = rSearchTmoS) AND ((rSearchTmoS - rSearchTmoS) = DL_WGE_Z)
        AND (rLostTmoS = rLostTmoS) AND ((rLostTmoS - rLostTmoS) = DL_WGE_Z)
        AND (rCenterTmoS = rCenterTmoS) AND ((rCenterTmoS - rCenterTmoS) = DL_WGE_Z);   // 九个浮点入参有限性 EN: the finiteness of all nine floating inputs
xParamBad := (NOT xFinAll) OR (rDeadbandMm < DL_WGE_Z) OR (rFindBandMm <= rDeadbandMm)
          OR (rMaxOffsetMm <= rFindBandMm) OR (rCorrRateMmS <= DL_WGE_Z) OR (rScanRateMmS <= DL_WGE_Z)
          OR (rSearchTmoS <= DL_WGE_Z) OR (rLostTmoS <= DL_WGE_Z) OR (rCenterTmoS <= DL_WGE_Z);   // 域闸与带间配比 EN: the domain gate and the band ordering
IF NOT xParamBad THEN                                                                              // 参数合法才换算 EN: convert only when the parameters are legal
    nMsSearch := REAL_TO_UDINT(rSearchTmoS * DL_WGE_K1000);                                        // 找边毫秒数 EN: the search milliseconds
    nMsLost := REAL_TO_UDINT(rLostTmoS * DL_WGE_K1000);                                            // 丢边毫秒数 EN: the lost milliseconds
    nMsCenter := REAL_TO_UDINT(rCenterTmoS * DL_WGE_K1000);                                        // 回中毫秒数 EN: the centering milliseconds
END_IF
xSensorUse := xSensorOk AND (NOT xParamBad);                                                       // 传感器可用判据 EN: the sensor usability test
rAbsOff := ABS(rEdgeOffsetMm);                                                                     // 偏移绝对值 [mm] EN: the offset magnitude

// 段2｜三只定时器 + 三只边沿实例无条件周期刷新（CASE 内不调用实例）
tonSearch(IN := (eState = E_DL_WebGuideState.EDGE_SEARCH), PT := UDINT_TO_TIME(nMsSearch));        // 找边计时 EN: the edge search timer
tonLost(IN := (eState = E_DL_WebGuideState.EDGE_LOST), PT := UDINT_TO_TIME(nMsLost));              // 丢边保持计时 EN: the edge lost timer
tonCenter(IN := (eState = E_DL_WebGuideState.CENTERING), PT := UDINT_TO_TIME(nMsCenter));          // 回中计时 EN: the centering timer
fbStartRise(CLK := xStart);                                                                        // 启动沿 EN: the start edge
fbStartFall(CLK := xStart);                                                                        // 复位沿 EN: the reset edge
fbRollRise(CLK := xRollChange);                                                                    // 换卷沿 EN: the roll change edge

// 段3｜输出预置（唯一预置点；EDGE_LOST 冻结语义在此体现为上拍快照）
rActCmdMmS := rLastCmd;                    // 指令预置为上拍快照（冻结保持） [mm/s] EN: preset the command to the previous snapshot
xMotionEnabled := FALSE;                   // 使能预置假 EN: preset the enable false
xFault := FALSE;                           // 故障标志预置假 EN: preset the fault flag false
nFaultCode := 0;                           // 故障码预置零 EN: preset the fault code to zero
nWarnCode := 0;                            // 信息码预置零 EN: preset the warning code to zero
xEdgeFound := (eState = E_DL_WebGuideState.TRACKING);   // 已找到边直映相态 EN: mirror the found state from the phase

// 段4｜全局安全闸：参数非法 / 运行中卷材缺失 → 锁故障；xStop 撤销指令回待机
IF xParamBad THEN
    nCodeLatch := DL_WGE_C_PARAM;                                                       // 参数非法锁存 EN: latch the parameter code
    xFault := TRUE;                                                                     // 置故障标志 EN: raise the fault flag
    nFaultCode := DL_WGE_C_PARAM;                                                       // 故障码出口 EN: publish the fault code
    eState := E_DL_WebGuideState.FAULT;                                                 // 迁故障相 EN: move to the fault phase
ELSIF (NOT xWebPresent) AND (eState <> E_DL_WebGuideState.IDLE) THEN
    nCodeLatch := DL_WGE_C_WEB;                                                         // 卷材缺失锁存 EN: latch the missing web code
    xFault := TRUE;                                                                     // 置故障标志 EN: raise the fault flag
    nFaultCode := DL_WGE_C_WEB;                                                         // 故障码出口 EN: publish the fault code
    eState := E_DL_WebGuideState.FAULT;                                                 // 迁故障相 EN: move to the fault phase
ELSIF xStop AND (eState <> E_DL_WebGuideState.IDLE) THEN
    rLastCmd := DL_WGE_Z;                                                               // 撤销型停车清空冻结快照，防止重启首拍陈指令 EN: a withdrawing stop clears the frozen snapshot so a restart cannot emit a stale command
    eState := E_DL_WebGuideState.IDLE;                                                  // 撤销型停车回待机 EN: a withdrawing stop returns to idle
END_IF

// 段5｜主状态机（ENUM + CASE，ELSE 兜底非法值）
IF eState <> E_DL_WebGuideState.FAULT THEN
CASE eState OF
E_DL_WebGuideState.IDLE:
    // 拍 N：待机；启动沿且卷材存在才进找边相（入相前置条件已含卷材与传感器）
    IF fbStartRise.Q AND xWebPresent AND (NOT xStop) AND xSensorUse THEN
        eState := E_DL_WebGuideState.EDGE_SEARCH;                                    // 本拍行为：进找边相 EN: enter the edge search phase
    END_IF

E_DL_WebGuideState.EDGE_SEARCH:
    // 拍 N：按偏移符号反方向扫描找边；进入判定带即进跟踪相，超时判 9601
    xMotionEnabled := TRUE;                                                          // 找边允许动作 EN: motion allowed for the search
    IF (NOT xSensorUse) THEN
        eState := E_DL_WebGuideState.EDGE_LOST;                                      // 本拍行为：传感器失效转丢边相 EN: the sensor failed, move to the lost phase
    ELSIF rAbsOff <= rFindBandMm THEN
        eState := E_DL_WebGuideState.TRACKING;                                       // 本拍行为：找到边进跟踪相 EN: the edge is found, enter tracking
    ELSIF tonSearch.Q THEN
        nCodeLatch := DL_WGE_C_SEARCH;                                               // 找边超时 EN: the edge search timed out
        xFault := TRUE;                                                              // 置故障标志 EN: raise the fault flag
        nFaultCode := DL_WGE_C_SEARCH;                                               // 故障码出口 EN: publish the fault code
        eState := E_DL_WebGuideState.FAULT;                                          // 迁故障相 EN: move to the fault phase
    ELSE
        IF rEdgeOffsetMm > DL_WGE_Z THEN                                             // 偏右则向左扫描 EN: scan left when the web sits right
            rCmd := -rScanRateMmS;                                                   // 负向扫描速度 [mm/s] EN: the negative scan velocity
        ELSE
            rCmd := rScanRateMmS;                                                    // 正向扫描速度 [mm/s] EN: the positive scan velocity
        END_IF
        rActCmdMmS := rCmd;                                                          // 落定本拍指令 [mm/s] EN: publish the command
        rLastCmd := rCmd;                                                            // 更新快照 [mm/s] EN: update the snapshot
    END_IF

E_DL_WebGuideState.TRACKING:
    // 拍 N：死区内不动、区外按偏移符号反方向纠偏；传感器失效转丢边相，偏移越限判参数类故障
    IF (NOT xSensorUse) THEN
        eState := E_DL_WebGuideState.EDGE_LOST;                                      // 本拍行为：丢边转保持相 EN: the edge is lost, move to the hold phase
    ELSIF fbRollRise.Q THEN
        eState := E_DL_WebGuideState.CENTERING;                                      // 本拍行为：换卷进回中相 EN: a roll change enters centering
    ELSIF rAbsOff > rMaxOffsetMm THEN
        nCodeLatch := DL_WGE_C_PARAM;                                                // 偏移越最大允许值，按参数/采样非法处理 EN: the offset exceeded the allowed maximum
        xFault := TRUE;                                                              // 置故障标志 EN: raise the fault flag
        nFaultCode := DL_WGE_C_PARAM;                                                // 故障码出口 EN: publish the fault code
        eState := E_DL_WebGuideState.FAULT;                                          // 迁故障相 EN: move to the fault phase
    ELSE
        xMotionEnabled := TRUE;                                                      // 跟踪允许动作 EN: motion allowed for tracking
        IF rAbsOff <= rDeadbandMm THEN                                               // 死区内不动 EN: no motion inside the dead band
            rCmd := DL_WGE_Z;                                                        // 指令给零 [mm/s] EN: give a zero command
        ELSIF rEdgeOffsetMm > DL_WGE_Z THEN                                          // 偏右则左移 EN: move left when the web sits right
            rCmd := -rCorrRateMmS;                                                   // 负向纠偏速度 [mm/s] EN: the negative correction velocity
        ELSE
            rCmd := rCorrRateMmS;                                                    // 正向纠偏速度 [mm/s] EN: the positive correction velocity
        END_IF
        rActCmdMmS := rCmd;                                                          // 落定本拍指令 [mm/s] EN: publish the command
        rLastCmd := rCmd;                                                            // 更新快照 [mm/s] EN: update the snapshot
    END_IF

E_DL_WebGuideState.EDGE_LOST:
    // 拍 N：丢边保持——使能保持并原样输出上一拍指令（真冻结，不是等效停车）；传感器恢复即回跟踪，保持超时判 9606
    // EN: hold on a lost edge, keeping the enable and republishing the previous command so the hold is a true freeze rather than an equivalent stop; recovery returns to tracking, a hold timeout raises 9606
    xMotionEnabled := TRUE;                                                          // 丢边保持仍维持使能 EN: keep the enable during the hold
    rActCmdMmS := rLastCmd;                                                          // 原样输出上一拍指令 [mm/s] EN: republish the previous command
    nWarnCode := DL_WGE_W_LOST;                                                      // 信息级：丢边保持中 EN: information class, the edge stays lost
    IF xSensorUse THEN
        eState := E_DL_WebGuideState.TRACKING;                                       // 本拍行为：传感器恢复回跟踪 EN: the sensor recovered, back to tracking
    ELSIF tonLost.Q THEN
        nCodeLatch := DL_WGE_C_LOST;                                                 // 丢边保持超时 EN: the edge lost hold timed out
        xFault := TRUE;                                                              // 置故障标志 EN: raise the fault flag
        nFaultCode := DL_WGE_C_LOST;                                                 // 故障码出口 EN: publish the fault code
        eState := E_DL_WebGuideState.FAULT;                                          // 迁故障相 EN: move to the fault phase
    END_IF

E_DL_WebGuideState.CENTERING:
    // 拍 N：换卷回中——按偏移缓慢回中，进死区即回跟踪，超时判 9603
    IF (NOT xSensorUse) THEN
        eState := E_DL_WebGuideState.EDGE_LOST;                                      // 本拍行为：传感器失效转丢边相 EN: the sensor failed, move to the lost phase
    ELSIF rAbsOff <= rDeadbandMm THEN
        eState := E_DL_WebGuideState.TRACKING;                                       // 本拍行为：回中完成进跟踪相 EN: centering done, enter tracking
    ELSIF tonCenter.Q THEN
        nCodeLatch := DL_WGE_C_CENTER;                                               // 回中超时 EN: the centering timed out
        xFault := TRUE;                                                              // 置故障标志 EN: raise the fault flag
        nFaultCode := DL_WGE_C_CENTER;                                               // 故障码出口 EN: publish the fault code
        eState := E_DL_WebGuideState.FAULT;                                          // 迁故障相 EN: move to the fault phase
    ELSE
        xMotionEnabled := TRUE;                                                      // 回中允许动作 EN: motion allowed for centering
        IF rEdgeOffsetMm > DL_WGE_Z THEN                                             // 偏右则左移 EN: move left when the web sits right
            rCmd := -rCorrRateMmS;                                                   // 负向回中速度 [mm/s] EN: the negative centering velocity
        ELSE
            rCmd := rCorrRateMmS;                                                    // 正向回中速度 [mm/s] EN: the positive centering velocity
        END_IF
        rActCmdMmS := rCmd;                                                          // 落定本拍指令 [mm/s] EN: publish the command
        rLastCmd := rCmd;                                                            // 更新快照 [mm/s] EN: update the snapshot
    END_IF

E_DL_WebGuideState.FAULT:
    // 故障相（本段被外层 IF 排除，保留分支以满足枚举穷举）
    xFault := TRUE;                                                                  // 保持故障标志 EN: keep the fault flag
    nFaultCode := nCodeLatch;                                                        // 锁存回放 EN: replay the latch

ELSE
    // 非法状态兜底：绝不停在未知相
    nCodeLatch := DL_WGE_C_PARAM;                                                    // 非法状态归参数码 EN: treat an illegal state as a parameter code
    xFault := TRUE;                                                                  // 置故障标志 EN: raise the fault flag
    nFaultCode := DL_WGE_C_PARAM;                                                    // 故障码出口 EN: publish the fault code
    eState := E_DL_WebGuideState.FAULT;                                              // 迁故障相 EN: move to the fault phase
END_CASE
END_IF

// 段6｜故障相锁存回放 + 复位沿（xStart 下降沿清除，复位后停 IDLE）
IF eState = E_DL_WebGuideState.FAULT THEN
    xFault := TRUE;                                                                  // 故障标志保持 EN: keep the fault flag
    nFaultCode := nCodeLatch;                                                        // 锁存回放，不按当下输入重推断 EN: replay the latch instead of re inferring
    nWarnCode := 0;                                                                  // 故障相不报信息级码 EN: no information class code in the fault phase
    xMotionEnabled := FALSE;                                                         // 撤销执行使能 EN: withdraw the motion enable
    rActCmdMmS := DL_WGE_Z;                                                          // 指令强制归零 [mm/s] EN: force the command to zero
    rLastCmd := DL_WGE_Z;                                                            // 快照归零，防复位后继承旧指令 [mm/s] EN: clear the snapshot so a reset cannot inherit a stale command
    IF fbStartFall.Q THEN
        nCodeLatch := 0;                                                             // 清除边：xStart 下降沿（头注释已声明） EN: clear on the falling edge of xStart
        eState := E_DL_WebGuideState.IDLE;                                           // 回待机 EN: back to idle
    END_IF
END_IF
END_FUNCTION_BLOCK

(* ---- FB_DL_WinderTensionTaperCtrl.st ---- *)
// FB_DL_WinderTensionTaperCtrl v1.0.0
(*==============================================================================
 * 功能描述: C4 收卷锥度张力控制。给定内圈张力 fTensionIn 与锥度系数 fTaperK，按当前
 *           卷径 fDiameter 外推张力设定（锥度模式）或恒张力模式，设定值经 fRampRate
 *           斜坡限速输出；模式切换与卷径突变均由斜坡自然平滑。卷径/张力限幅与组态
 *           非法、非有限输入防御齐备。
 * 接口契约: 输入 bEnable/eModeReq/fTensionIn/fTaperK/fDiameter/fDiaMin/fDiaMax/
 *           fTensionMin/fTensionMax/fRampRate/fDtSec/bReset；
 *           输出 fTensionSet/eModeAct/bValid/eState/bError/nErrId。
 * 边界: ① 组态闸：fDiaMin<=0、fDiaMax<fDiaMin、fTensionMin<0、fTensionMax<=fTensionMin、
 *           fRampRate<=0、fDtSec<=0 或任一浮点引脚 NaN → 故障锁存；② 卷径先钳位到
 *           [fDiaMin,fDiaMax] 再进锥度外推（R4 防越界）；③ 一枚 R_TRIG 段 0 无条件刷新；
 *           ④ 零全局耦合。
 * 码表: 16#0007_0302 故障级总码（组态非法/非有限输入/非法相位，锁存至 bReset 上升沿）。
 * 修订历史: 2026-11-23  v1.0.0  R74 首版
 *==============================================================================*)

TYPE E_DL_WttMode :
(
    eConstant := 0,   // 恒张力模式（不随卷径外推）/ Constant tension mode
    eTaper    := 1    // 锥度张力模式（随卷径线性外推）/ Taper tension mode
);
END_TYPE

TYPE E_DL_WttState :
(
    eIdle  := 0,      // 待机（设定值冻结保持）/ Idle, setpoint frozen
    eRun   := 10,     // 运行（斜坡跟随目标）/ Running, ramp toward target
    eFault := 90      // 故障锁存相（仅复位沿迁出）/ Fault latched, exit by reset edge only
);
END_TYPE

FUNCTION_BLOCK FB_DL_WinderTensionTaperCtrl
VAR_INPUT
    bEnable     : BOOL := FALSE;         // 使能（FALSE 冻结输出保持）[-] / Enable, FALSE freezes output
    eModeReq    : E_DL_WttMode := E_DL_WttMode.eTaper;   // 张力模式请求 [枚举] / Tension mode request
    fTensionIn  : REAL := 50.0;          // 内圈张力给定，域 > 0 [N] / Inner tension setpoint [N]
    fTaperK     : REAL := 0.0005;        // 锥度系数，域 >= 0 [1/mm] / Taper coefficient [1/mm]
    fDiameter   : REAL := 100.0;         // 当前卷径反馈 [mm] / Current roll diameter [mm]
    fDiaMin     : REAL := 100.0;         // 卷径下限（纸芯径），域 > 0 [mm] / Minimum diameter [mm]
    fDiaMax     : REAL := 800.0;         // 卷径上限，域 >= fDiaMin [mm] / Maximum diameter [mm]
    fTensionMin : REAL := 0.0;           // 张力下限，域 >= 0 [N] / Tension lower limit [N]
    fTensionMax : REAL := 200.0;         // 张力上限，域 > fTensionMin [N] / Tension upper limit [N]
    fRampRate   : REAL := 10.0;          // 设定值斜坡速率，域 > 0 [N/s] / Ramp rate [N/s]
    fDtSec      : REAL := 0.010;         // 任务周期 [s]，域 > 0 / Task period [s], domain > 0
    bReset      : BOOL := FALSE;         // 复位，上升沿清故障锁存 [-] / Reset edge clears fault
END_VAR
VAR_OUTPUT
    fTensionSet : REAL := 0.0;           // 张力设定输出（斜坡后，限幅内）[N] / Tension setpoint output [N]
    eModeAct    : E_DL_WttMode;          // 当前生效模式出口 [枚举] / Active mode outlet
    bValid      : BOOL;                  // 设定值有效回执 [-] / Setpoint validity receipt
    eState      : E_DL_WttState;         // 状态出口，段尾单点映射 / State outlet
    bError      : BOOL;                  // 故障锁存标志 [-] / Fault latch flag
    nErrId      : UDINT;                 // 事件码，0 = 无事件 / Event code, 0 = none
END_VAR
VAR
    _eState    : E_DL_WttState := E_DL_WttState.eIdle;   // 内部相位（CASE 唯一写入目标） / Internal phase
    rtReset    : R_TRIG;                 // 复位沿实例，段 0 无条件刷新 / Reset edge instance
    _fTarget   : REAL := 0.0;            // 本拍目标张力（限幅后）[N] / Target tension this scan [N]
    _fSetInt   : REAL := 0.0;            // 内部斜坡设定值（锁存量）[N] / Internal ramped setpoint
    _fDiaEff   : REAL := 0.0;            // 钳位后有效卷径 [mm] / Clamped effective diameter [mm]
    _fStep     : REAL := 0.0;            // 本拍斜坡步长 [N] / Ramp step this scan
    _bCfgBad   : BOOL;                   // 组态非法当拍量 [-] / Illegal configuration this scan
    _bNonFin   : BOOL;                   // 输入非有限当拍量 [-] / Non-finite input this scan
    _bFault    : BOOL;                   // 故障锁存位（锁存量） / Latched fault bit
    _uFault    : UDINT;                  // 故障码锁存（锁存量） / Latched fault code
    _eModeInt  : E_DL_WttMode := E_DL_WttMode.eTaper;    // 生效模式锁存 / Active mode latch
END_VAR

(* —— 段 0：沿实例无条件周期刷新 —— *)
rtReset(CLK := bReset);                                            // 复位沿，每拍必调 / Reset edge, called every scan

(* —— 段 1：单拍量预清零（锁存量 _fSetInt/_eModeInt/_bFault/_uFault 不入清单） —— *)
bValid := FALSE;                                                   // 有效回执预清（运行相回填） / Validity preset
bError := FALSE;                                                   // 故障标志预清（置位处同拍回填） / Error flag preset
nErrId := 16#0000_0000;                                            // 事件码缺省无事件 / Event code default none

(* —— 段 2：组态域闸与非有限闸（覆盖全部参与引脚） —— *)
_bNonFin := (fTensionIn <> fTensionIn) OR (fTaperK <> fTaperK)     // 给定与系数 NaN 自反判 / NaN self-reflexive tests
         OR (fDiameter <> fDiameter) OR (fDiaMin <> fDiaMin)       // 卷径引脚 NaN 判 / Diameter NaN tests
         OR (fDiaMax <> fDiaMax) OR (fTensionMin <> fTensionMin)   // 限幅引脚 NaN 判 / Limit NaN tests
         OR (fTensionMax <> fTensionMax) OR (fRampRate <> fRampRate)// 上限与速率 NaN 判 / Upper limit and rate NaN tests
         OR (fDtSec <> fDtSec);                                    // 周期 NaN 判 / Period NaN test
_bCfgBad := (fDiaMin <= 0.0) OR (fDiaMax < fDiaMin)                // 卷径域闸 / Diameter domain gates
         OR (fTensionMin < 0.0) OR (fTensionMax <= fTensionMin)    // 张力限幅域闸 / Tension limit gates
         OR (fRampRate <= 0.0) OR (fDtSec <= 0.0)                  // 速率与周期域闸 / Rate and period gates
         OR (fTensionIn <= 0.0);                                   // 给定正值闸 / Positive setpoint gate

(* —— 段 3：故障锁存与解除（R45 配对；解除式全当拍量） —— *)
IF _bCfgBad THEN                                                   // 组态非法 / Illegal configuration
    _uFault := 16#0007_0302;                                       // 故障级总码 / Fault-level code
    _bFault := TRUE;
    bError  := TRUE;
END_IF
IF (NOT _bFault) AND _bNonFin THEN                                 // 输入非有限 / Non-finite input
    _uFault := 16#0007_0302;
    _bFault := TRUE;
    bError  := TRUE;
END_IF
IF rtReset.Q AND (NOT _bCfgBad) AND (NOT _bNonFin) THEN            // 解除沿（当拍量） / Release edge
    _bFault := FALSE;                                              // 清故障锁存 / Clear fault latch
    _uFault := 16#0000_0000;                                       // 清故障码 / Clear fault code
    IF _eState = E_DL_WttState.eFault THEN
        _eState := E_DL_WttState.eIdle;                            // 故障相唯一迁出路径 / Sole exit from fault phase
    END_IF
END_IF

(* —— 段 4：相位机（ENUM 全成员显式标签 + ELSE 兜底） —— *)
CASE _eState OF

E_DL_WttState.eIdle:
    IF (NOT _bFault) AND bEnable THEN                              // 出口 1：使能进运行 / Enable enters run
        _eModeInt := eModeReq;                                     // 锁存生效模式 / Latch active mode
        _eState := E_DL_WttState.eRun;
    ELSIF _bFault THEN                                             // 出口 2：故障锁存 / Fault latched
        _eState := E_DL_WttState.eFault;
    END_IF

E_DL_WttState.eRun:
    IF (NOT bEnable) THEN                                          // 出口 1：撤使能回待机（设定值冻结保持） / Disable, setpoint frozen
        _eState := E_DL_WttState.eIdle;
    ELSIF _bFault THEN                                             // 出口 2：故障锁存 / Fault latched
        _eState := E_DL_WttState.eFault;
    ELSE
        _eModeInt := eModeReq;                                     // 模式请求每拍跟随（切换由斜坡平滑） / Mode follows request, ramp smooths
        _fDiaEff := fDiameter;                                     // 卷径预装 / Diameter preloaded
        IF _fDiaEff < fDiaMin THEN                                 // 卷径下限钳位（R4 防越界） / Clamp to lower bound
            _fDiaEff := fDiaMin;
        END_IF
        IF _fDiaEff > fDiaMax THEN                                 // 卷径上限钳位 / Clamp to upper bound
            _fDiaEff := fDiaMax;
        END_IF
        IF _eModeInt = E_DL_WttMode.eTaper THEN                    // 锥度模式：按卷径线性外推 / Taper mode, linear extrapolation
            _fTarget := fTensionIn * (1.0 + fTaperK * (_fDiaEff - fDiaMin));   // 锥度外推 [N] / Taper extrapolation
        ELSE                                                       // 恒张力模式 / Constant mode
            _fTarget := fTensionIn;                                // 目标 = 给定 / Target equals setpoint
        END_IF
        IF _fTarget < fTensionMin THEN                             // 张力下限饱和钳位 / Saturate at lower limit
            _fTarget := fTensionMin;
        END_IF
        IF _fTarget > fTensionMax THEN                             // 张力上限饱和钳位 / Saturate at upper limit
            _fTarget := fTensionMax;
        END_IF
        _fStep := fRampRate * fDtSec;                              // 本拍斜坡步长 [N] / Ramp step this scan
        IF _fSetInt < (_fTarget - _fStep) THEN                     // 上升斜坡限速 / Upward ramp limited
            _fSetInt := _fSetInt + _fStep;
        ELSIF _fSetInt > (_fTarget + _fStep) THEN                  // 下降斜坡限速 / Downward ramp limited
            _fSetInt := _fSetInt - _fStep;
        ELSE
            _fSetInt := _fTarget;                                  // 步长内直达目标 / Within step, reach target
        END_IF
    END_IF

E_DL_WttState.eFault:
    ;                                                              // 故障相：仅段 3 复位沿可迁出 / Only the reset edge leaves this phase

ELSE
    _uFault := 16#0007_0302;                                       // 故障级：非法相位兜底 / Illegal-phase fallback
    _bFault := TRUE;
    bError  := TRUE;
    _eState := E_DL_WttState.eFault;                               // 强拉故障相 / Force fault phase

END_CASE

(* —— 段 5：出口单点映射（名实同源；锁存码回放；故障相安全侧） —— *)
IF (_eState = E_DL_WttState.eRun) AND (NOT _bFault) THEN
    fTensionSet := _fSetInt;                                       // 运行相输出斜坡设定 / Run phase outputs ramped setpoint
    bValid := TRUE;                                                // 有效回执 / Validity receipt
END_IF
eModeAct := _eModeInt;                                             // 模式出口 / Mode outlet
IF _bFault THEN
    fTensionSet := fTensionMin;                                    // 故障相安全侧：输出张力下限 / Safe side in fault
    nErrId := _uFault;                                             // 故障锁存码回放 / Replay latched fault code
END_IF
bError := _bFault;                                                 // 故障标志与锁存同源 / Flag from latch
eState := _eState;                                                 // 状态出口 / State outlet

END_FUNCTION_BLOCK

(* ---- FB_DL_WindingAlignEdge.st ---- *)
//==============================================================================
// 功能块：FB_DL_WindingAlignEdge ｜ 中文名称：卷绕极片边缘跟随与蛇形抑制
// 所属子库：DL_Motion ｜ 版本：v1.0.0 ｜ 兼容：CODESYS V3.5+ / TwinCAT 3 / 汇川 InoProShop
// 功能描述：极片边缘跟随纠偏——边缘传感器上升沿锁存轴位置为边缘基准，
//           偏差 = 锁存边缘 - 目标边缘，经一阶低通滤波（alpha 加权，滤
//           高频毛刺）与每拍步进限幅（蛇形抑制：禁止纠偏输出大幅摆动）
//           后乘增益输出纠偏百分比；纠偏输出受行程窗口拦截（超限钳位
//           + 信息提示）。相邻边沿间轴位移超过物理上限判传感器跳变/
//           双沿，锁存故障（防假边缘基准污染纠偏链）。
// 遗留假设（R95 代理阈值三句）：① 代理值 = fCycleTimeS 组态扫描周期
//           [秒]（步进限幅的换算基量）；② 覆盖 0.001~0.1 秒任务周期
//           范围；③ 覆盖不到的区间由调用方按实际任务周期重设该引脚
//           负责，该假设挂编译验证债。
// 开源溯源 (Origin)：道莅原创实现（参考卷绕纠偏（边缘跟随）工程惯例 分类与参数域）
// 单位表：轴位置[毫米] / 边缘目标[毫米] / 传感器偏置[毫米] / 偏差[毫米] /
//         增益[百分数每毫米] / 行程限[毫米] / 跳变限[毫米] / 增益系数[无量纲]
// 错误码表：16#0004_01E5 信息级（边缘锁存更新：新边沿被锁存为基准，不置
//           bError）/ 16#0004_01E6 信息级（纠偏输出达行程限幅，不置
//           bError）/ 16#0004_0303 故障级（组态非法：增益系数/行程限/
//           跳变限域、周期 <= 0 或任一输入非有限，置 bError）/
//           16#0004_0304 故障级（边沿跳变超物理上限：相邻边沿间轴位移
//           超 fMaxJumpMm，判传感器跳变/双沿，锁存故障，置 bError——
//           该场景不可由 0303 的组态类判据观测，属运行信号独立域）/
//           16#0004_0305 故障级兜底（状态机落 ELSE，置 bError）
// 状态机：E_DL_WindAlignState（四态：eIdle=0 / eFollow=10 / eFault=99），
//           实际为三态，CASE 含 ELSE 兜底，ELSE 置 0305 并冻结输出零
// 边界行为：① 组态非法 → 故障态锁存，bReset 复位；② 未锁存边缘前
//           纠偏输出保持 0（无基准不放行）；③ 滤波系数域 [0, 1]，= 0
//           即冻结滤波值（等于不更新）；④ 纠偏输出钳 +/- 行程限 + 信息
//           01E6；⑤ 未使能输出冻结零并 bValid := FALSE（锁存基准保持，
//           复能即续走）；⑥ 安全侧 = 跳变故障冻结纠偏输出为 0，禁止
//           假基准驱动机构。
// 修订历史：v1.0.0 2026-11-17 首版（R24 派单 · ROADMAP P1 §806）
//==============================================================================

(*------------------------------------------------------------------------------
 * 枚举: E_DL_WindAlignState（归属本功能块，同文件发布，全库唯一定义）
 * 含义: 边缘跟随相位，每个成员在 CASE 中有且仅有一个标签。
 *-----------------------------------------------------------------------------*)
TYPE E_DL_WindAlignState :
(
    eIdle   := 0,   // 空闲：未使能 / Idle, not enabled
    eFollow := 10,  // 跟随：纠偏闭环运行 / Follow, correction loop running
    eFault  := 99   // 故障：组态非法/边沿跳变/非法状态 / Fault, config, edge jump or illegal state
);
END_TYPE

FUNCTION_BLOCK FB_DL_WindingAlignEdge
VAR_INPUT
    bEnable       : BOOL;                   // 跟随使能 [—] / Follow enable
    bReset        : BOOL;                   // 故障复位 [—]，上升沿清锁存 / Fault reset, rising edge clears latches
    bEdgeSensor   : BOOL;                   // 边缘传感器电平 [—]（TRUE = 检出极片边缘） / Edge sensor level, TRUE on the edge
    fAxisPosMm    : LREAL;                  // 轴位置实测 [毫米]（纠偏机构位置基准） / Axis position [mm]
    fTargetEdgeMm : LREAL := 0.0;           // 目标边缘位置 [毫米] / Target edge position [mm]
    fSensorOffsetMm : LREAL := 0.0;         // 传感器安装偏置 [毫米]（锁存值补偿） / Sensor mounting offset [mm]
    fFilterAlpha  : LREAL := 0.2;           // 一阶滤波系数 [无量纲]，域 [0, 1]，0 = 冻结滤波值 / First-order filter alpha, domain 0..1
    fGainPctPerMm : LREAL := 10.0;          // 纠偏增益 [百分数每毫米] / Correction gain [percent/mm]
    fTravelLimitMm: LREAL := 20.0;          // 纠偏行程限 [毫米]，须 > 0 / Correction travel limit [mm], must be > 0
    fMaxJumpMm    : LREAL := 5.0;           // 相邻边沿位移物理上限 [毫米]，须 > 0 / Max inter-edge displacement [mm], must be > 0
    fCycleTimeS   : LREAL := 0.01;          // 任务扫描周期 [秒]，须 > 0（R95 代理阈值） / Task scan cycle [s], must be > 0, R95 proxy
END_VAR
VAR_OUTPUT
    fCorrectOutPct : LREAL;                 // 纠偏输出 [百分数]，-100..100，行程限内 / Correction output [percent], within the travel limit
    fOffsetMm      : LREAL;                 // 滤波后边缘偏差 [毫米]（诊断出口） / Filtered edge offset [mm], diagnostics outlet
    bEdgeLatch     : BOOL;                  // 边缘锁存有效 [—] / Edge latch valid
    eState         : E_DL_WindAlignState;   // 相位出口 [—] / Phase outlet
    eErr           : UDINT;                 // 错误码，0 = 无错，码位 16#0004_01E5 起信息级、16#0004_0303 起故障级（分带见错误码表） / Error code, 0 = no error, band info/fault per the code table
    bError         : BOOL;                  // 故障级标志，仅故障级错误置位 / Fault-class flag, set only on fault-level codes
    bValid         : BOOL;                  // 输出可用标志 / Outputs usable flag
END_VAR
VAR
    fbEdge    : R_TRIG;                     // 边缘沿检测（待机/故障分支同样无条件刷新） / Edge detector, refreshed unconditionally
    _eState   : E_DL_WindAlignState := E_DL_WindAlignState.eIdle; // 当前相位 / Current phase
    _bCfgBad  : BOOL;                       // 组态非法锁存 / Illegal config latch
    _bJumpBad : BOOL;                       // 边沿跳变锁存 / Edge jump fault latch
    _bInfoLatch: BOOL;                      // 锁存更新信息当拍标志 / Latch-update info flag of this scan
    _bInfoClip: BOOL;                       // 限幅信息当拍标志 / Clamp info flag of this scan
    _fEdgeCap : LREAL;                      // 锁存边缘基准 [毫米] / Latched edge reference [mm]
    _fEdgePrev: LREAL;                      // 上次锁存边缘基准 [毫米]（跳变判据基准） / Previous latched edge [mm]
    _fOffFilt : LREAL;                      // 滤波后偏差内部量 [毫米] / Filtered offset internal [mm]
    _fOutPrev : LREAL;                      // 上拍纠偏输出快照 [百分数]（步进限幅基准） / Previous-scan correction snapshot [percent]
    _bHaveL   : BOOL;                       // 已锁存标志 / Latch-present flag
    _bIllegal : BOOL;                       // 非法状态标志 / Illegal state flag
    _bInit    : BOOL := FALSE;              // 首扫标志，初值 FALSE 取非判定 / First-scan flag, tested negated
END_VAR
VAR CONSTANT
    DL_WAE_INF     : LREAL := 1.7976931348623157E308; // LREAL 幅值上限 / LREAL magnitude ceiling
    DL_WAE_EPS     : LREAL := 1.0E-6;       // 浮点判零容差 [毫米] / Float zero tolerance [mm]
    DL_WAE_SLEW_PCTS: LREAL := 50.0;        // 纠偏最大变化率 [百分数每秒]（蛇形抑制硬限） / Max correction slew rate [percent/s]
    DL_WAE_OUT_MAX : LREAL := 100.0;        // 纠偏输出满幅 [百分数] / Correction full scale [percent]
    DL_WAE_ZERO    : LREAL := 0.0;          // 零值常量，避免裸字面量 [混合] / Zero constant, avoids a bare literal
    DL_WAE_ONE     : LREAL := 1.0;          // 单位常量 [无量纲] / Unity constant
END_VAR

(*------------------------------------------------------------------------------
 * 段 1｜每拍预置：纠偏输出先清（安全侧），单拍标志预清零
 *      Correction cleared fail-safe first, one-shot flags pre-cleared
 *-----------------------------------------------------------------------------*)
fCorrectOutPct := DL_WAE_ZERO;           // 纠偏输出先清（跟随态在段 5 重置） / Correction cleared first
fOffsetMm := DL_WAE_ZERO;                // 偏差出口每拍重算 / Offset outlet recomputed
eErr   := 16#0000_0000;                  // 错误码每拍重算 / Error code recomputed
bError := FALSE;                         // 故障标志每拍重算 / Fault flag recomputed
bValid := FALSE;                         // 可用标志每拍重算 / Usable flag recomputed
_bInfoLatch := FALSE;                    // 锁存信息预清零 / Latch info pre-cleared
_bInfoClip  := FALSE;                    // 限幅信息预清零 / Clamp info pre-cleared
_bIllegal   := FALSE;                    // 非法状态预清零 / Illegal flag pre-cleared

(*------------------------------------------------------------------------------
 * 段 2｜首扫初始化
 *      First-scan initialisation
 *-----------------------------------------------------------------------------*)
IF NOT _bInit THEN
    _eState   := E_DL_WindAlignState.eIdle; // 相位空闲起步 / Phase starts idle
    _bCfgBad  := FALSE;                  // 组态锁存清零 / Config latch cleared
    _bJumpBad := FALSE;                  // 跳变锁存清零 / Jump latch cleared
    _bHaveL   := FALSE;                  // 锁存标志清零 / Latch flag cleared
    _fOffFilt := DL_WAE_ZERO;            // 滤波值从零起步 / Filter starts at zero
    _fOutPrev := DL_WAE_ZERO;            // 输出快照从零起步 / Output snapshot starts at zero
    _bInit    := TRUE;                   // 首扫只做一次 / The first scan runs once
END_IF

(*------------------------------------------------------------------------------
 * 段 3｜组态防御闸：非有限（R79）+ 增益/行程/跳变/周期域
 *      Configuration defense gates
 *-----------------------------------------------------------------------------*)
IF (fAxisPosMm <> fAxisPosMm) OR (ABS(fAxisPosMm) > DL_WAE_INF)
   OR (fFilterAlpha <> fFilterAlpha) OR (ABS(fFilterAlpha) > DL_WAE_INF)
   OR (fGainPctPerMm <> fGainPctPerMm) OR (ABS(fGainPctPerMm) > DL_WAE_INF)
   OR (fTravelLimitMm <> fTravelLimitMm) OR (ABS(fTravelLimitMm) > DL_WAE_INF)
   OR (fMaxJumpMm <> fMaxJumpMm) OR (ABS(fMaxJumpMm) > DL_WAE_INF)
   OR (fCycleTimeS <> fCycleTimeS) OR (ABS(fCycleTimeS) > DL_WAE_INF) THEN
    _bCfgBad := TRUE;                    // 非有限归组态非法锁存 / Non-finite folded into the config latch
END_IF
IF (NOT _bCfgBad) AND ((fFilterAlpha < DL_WAE_ZERO) OR (fFilterAlpha > DL_WAE_ONE)
   OR (fTravelLimitMm <= DL_WAE_EPS) OR (fMaxJumpMm <= DL_WAE_EPS)
   OR (fCycleTimeS <= DL_WAE_EPS)) THEN
    _bCfgBad := TRUE;                    // 增益系数/行程限/跳变限/周期域非法锁存 / Gain, travel, jump and cycle domains latched
END_IF
IF bReset THEN
    _bCfgBad  := FALSE;                  // 复位清组态锁存 / Reset clears the config latch
    _bJumpBad := FALSE;                  // 复位清跳变锁存 / Reset clears the jump latch
END_IF

(*------------------------------------------------------------------------------
 * 段 4｜边缘沿检测无条件刷新（R40：CASE 之外每拍必调）
 *      Edge detection refreshed unconditionally per R40
 *-----------------------------------------------------------------------------*)
fbEdge(CLK := bEdgeSensor);              // 边缘沿检测 / Edge detection

(*------------------------------------------------------------------------------
 * 段 5｜相位机与纠偏链（CASE 含 ELSE 兜底；未使能/异常落故障态）
 *      Phase machine and the correction chain
 *-----------------------------------------------------------------------------*)
IF (NOT bEnable) OR _bCfgBad OR _bJumpBad THEN
    _eState := E_DL_WindAlignState.eFault; // 未使能或异常转故障态（输出零） / Not enabled or anomaly, fault, output zero
ELSE
CASE _eState OF

    E_DL_WindAlignState.eIdle:             // 空闲：使能进跟随（基准未锁存则输出保持零）
        IF bEnable THEN
            _eState := E_DL_WindAlignState.eFollow; // 进跟随 / To follow
        END_IF

    E_DL_WindAlignState.eFollow:           // 跟随：沿锁存 + 滤波 + 步进限幅 + 行程拦截
        IF NOT bEnable THEN
            _eState := E_DL_WindAlignState.eFault; // 使能撤销转故障 / Enable dropped, fault
        END_IF
        IF fbEdge.Q THEN                   // 新边沿：跳变校验通过才锁存（R80 三段式）
            IF _bHaveL AND (ABS(fAxisPosMm - _fEdgePrev) > fMaxJumpMm) THEN
                _bJumpBad := TRUE;         // 相邻边沿位移超物理上限（拍 N 进入） / Inter-edge displacement beyond the physical limit
                _eState := E_DL_WindAlignState.eFault; // 本拍转出：进故障冻结 / To fault, frozen
            ELSE
                _fEdgeCap := fAxisPosMm - fSensorOffsetMm; // 锁存边缘基准（含安装偏置补偿） [毫米] / Latch the edge with offset compensation
                _fEdgePrev := _fEdgeCap;   // 跳变判据基准推进 / Jump-reference advanced
                _bHaveL := TRUE;           // 锁存有效 / Latch valid
                _bInfoLatch := TRUE;       // 锁存更新提示（信息级） / Latch-update notice, info
            END_IF
        END_IF
        IF (_eState = E_DL_WindAlignState.eFollow) AND _bHaveL THEN
            fOffsetMm := _fEdgeCap - fTargetEdgeMm; // 原始偏差 [毫米] / Raw offset [mm]
            _fOffFilt := _fOffFilt + fFilterAlpha * (fOffsetMm - _fOffFilt); // 一阶低通滤波 [毫米] / First-order low-pass filter
            fOffsetMm := _fOffFilt;        // 滤波后偏差出口 / Filtered offset outlet
            fCorrectOutPct := fGainPctPerMm * _fOffFilt; // 增益映射 [百分数] / Gain mapping
            fCorrectOutPct := MIN(MAX(fCorrectOutPct,
                _fOutPrev - DL_WAE_SLEW_PCTS * fCycleTimeS),
                 _fOutPrev + DL_WAE_SLEW_PCTS * fCycleTimeS); // 每拍步进限幅（蛇形抑制：变化率受限） / Per-scan slew clamp, anti-serpentine
            fCorrectOutPct := MIN(MAX(fCorrectOutPct,
                -MIN(fTravelLimitMm * fGainPctPerMm, DL_WAE_OUT_MAX),
                 MIN(fTravelLimitMm * fGainPctPerMm, DL_WAE_OUT_MAX))); // 行程窗拦截钳位（变化率限后二次钳位） / Travel-window clamp after the slew
            IF ABS(fCorrectOutPct) >= (MIN(fTravelLimitMm * fGainPctPerMm, DL_WAE_OUT_MAX) - DL_WAE_EPS) THEN
                _bInfoClip := TRUE;        // 达行程限幅提示（信息级） / Travel-limit notice, info
            END_IF
            _fOutPrev := fCorrectOutPct;   // 上拍输出快照推进（步进限幅基准） / Previous-output snapshot advanced
        END_IF

    E_DL_WindAlignState.eFault:            // 故障：复位沿且原因消失回空闲
        IF bReset AND (NOT _bCfgBad) AND (NOT _bJumpBad) THEN
            _eState := E_DL_WindAlignState.eIdle; // 回空闲 / Back to idle
        END_IF

    ELSE                                   // 非法状态兜底（R21：CASE 必带 ELSE）
        _bIllegal := TRUE;                 // 标记非法状态 / Flag the illegal state
        fCorrectOutPct := DL_WAE_ZERO;     // 输出冻结零（安全侧） / Output frozen at zero
        _eState := E_DL_WindAlignState.eFault; // 回故障态 / Back to fault
END_CASE
END_IF

(*------------------------------------------------------------------------------
 * 段 6｜码位出口与放行（故障级码 3 行内置 bError，R45/R101 配对）
 *      Code outlet and release, fault codes paired with bError
 *-----------------------------------------------------------------------------*)
IF _bIllegal THEN
    eErr   := 16#0004_0305;                // 故障级：状态机兜底 / Fault: state machine fallback
    bError := TRUE;                        // 置故障标志 / Raise the fault flag
ELSIF _bJumpBad THEN
    eErr   := 16#0004_0304;                // 故障级：边沿跳变超物理上限 / Fault: edge jump beyond the physical limit
    bError := TRUE;                        // 置故障标志 / Raise the fault flag
ELSIF _bCfgBad THEN
    eErr   := 16#0004_0303;                // 故障级：组态非法 / Fault: illegal configuration
    bError := TRUE;                        // 置故障标志 / Raise the fault flag
ELSIF _bInfoClip THEN
    eErr := 16#0004_01E6;                  // 信息级：纠偏输出达行程限幅 / Info: correction at the travel limit
ELSIF _bInfoLatch THEN
    eErr := 16#0004_01E5;                  // 信息级：边缘锁存更新 / Info: edge latch updated
END_IF

bEdgeLatch := _bHaveL AND (NOT bError);  // 锁存有效出口（故障时不放行） / Latch-valid outlet, gated in fault
bValid := (NOT bError) AND bEnable AND (_eState = E_DL_WindAlignState.eFollow); // 仅跟随态放行 / Usable only in the follow phase
eState := _eState;                       // 相位出口 / Phase outlet
END_FUNCTION_BLOCK

(* ---- FB_DL_WindingLayerCounter.st ---- *)
(*
    FB_DL_WindingLayerCounter —— 卷绕层数计数
    ------------------------------------------------------------------
    分类      : DL_Motion / Winding
    前缀      : FB_DL_
    版本      : 1.0.0
    溯源      : 层数递推为公开几何关系（层数 = (卷径 − 芯径) / (2·厚度)）；
                与算直径件构成「算一个值 / 数一件事」的职责切分；
                交叉校核、饱和钳位、换卷语义、错误分级与码位 100% 自有；
                clean-room 重写，未复制任何闭源厂商源码
    平台      : 纯 IEC 61131-3，CODESYS V3.5+ / TwinCAT 3 / InoProShop 通用
    作者      : 道莅代码库 · PLC编程专家（R19）
    ------------------------------------------------------------------
    功能说明  : 由「卷径 + 芯径 + 材料厚度」推算已绕层数与剩余层数，并与卷轴累计圈计数
                交叉校核：两者差超过 1 层即置 bInconsistent，但只提示不报故障——
                打滑/叠绕/测距噪声在薄膜与极片卷绕里是常态，报故障会误停整条线。
                核心防御：① 厚度或芯径非法即故障级 02E7 并冻结层数（厚度在分母上，
                   是本件除零唯一出口）；
                ② 卷径小于芯径即故障级 02E8——物理上不可能，通常是测距件故障或
                   参数填反，此时硬算会得到负层数；
                ③ 层数超上限只钳位并置信息码；④ 剩余层数由上限减去已绕层数，下溢钳 0；
                ⑤ 等效厚度反推的分母用 MAX(|圈数|, 1) 而不是除零闸——圈数为 0 是开机常态；
                ⑥ 圈计数取模长参与校核（层数是标量，方向由 bDirPositive 另行表达），
                   取模长先升位到 LINT 再取负，规避 DINT 最小值取负回绕（R55）。
                职责边界：卷径测量与滤波归测距/卷径件，本件只数层；张力与排线另有专件。
    错误码    : 16#0004_01D3 层数超上限已钳位 / 圈计数与卷径推算不一致（打滑或叠绕，仅提示）——信息级，正常防御
                16#0004_01D4 预留禁用（信息级，不得挪用）
                16#0004_02E7 厚度或芯径非法（<= 0 / 非有限）——故障级，层数冻结
                16#0004_02E8 卷径非有限或小于芯径（含测距件故障）——故障级，层数冻结
                16#0004_02E9 预留禁用（故障级，不得挪用）
    码位总账  : 16#0004_01D3 用 / 16#0004_01D4 预留 ｜ 16#0004_02E7 用 / 16#0004_02E8 用 / 16#0004_02E9 预留
    状态机    : R6 标注 N/A —— 本组件为纯函数无顺序状态机，无 CASE 可写，非法状态不可能出现
    采样约定  : fbTrigReset / fbTrigNewRoll 在本体首部无条件刷新；本件无时间量，
                bLayerEdge 为单周期脉冲（每拍先清后置），结论与任务周期无关。
    修订记录  : 2026-11-16 v1.0.0 首次入库（R19）
*)
FUNCTION_BLOCK FB_DL_WindingLayerCounter
VAR_INPUT
    bEnable         : BOOL;                   // 使能，FALSE 冻结层数 / enable, FALSE freezes the layer count
    bReset          : BOOL;                   // 复位，上升沿清零（含累计统计）/ reset, rising edge clears everything including the statistics
    bNewRoll        : BOOL;                   // 换卷，上升沿视为换卷（保留累计统计）/ new roll, rising edge starts a new roll while keeping the statistics
    fCoilDiameter   : REAL := 76.2;           // 当前卷径（外部卷径件/测距给出）[mm] / current coil diameter from the measurement block [mm]
    fCoreDiameter   : REAL := 76.2;           // 芯径 [mm]，必须 > 0 / core diameter [mm], must be > 0
    fThickness      : REAL := 0.1;            // 材料厚度（含隔膜/铜箔）[mm]，必须 > 0 / material thickness [mm], must be > 0
    diRevCount      : DINT := 0;              // 卷轴累计圈计数（方向敏感）[圈] / accumulated shaft revolutions, direction sensitive [rev]
    uLayerMax       : UINT := 5000;           // 层数饱和上限 [层]，范围 10~60000 / layer saturation bound [layer], range 10~60000
    bDirPositive    : BOOL := TRUE;           // 当前旋转方向（反向时圈计数按模长校核）/ current rotation direction, magnitude is used for the cross-check
END_VAR
VAR_OUTPUT
    uLayerDone      : UINT;                   // 已绕层数（由卷径推算）[层] / layers wound, derived from the diameter [layer]
    uLayerRemain    : UINT;                   // 剩余层数（相对上限）[层] / remaining layers relative to the bound [layer]
    bLayerEdge      : BOOL;                   // 层数变化单周期脉冲 / single-cycle pulse on a layer change
    bInconsistent   : BOOL;                   // 圈计数与卷径推算不一致（超过 1 层）/ the revolution count disagrees with the diameter estimate by more than one layer
    fThicknessEst   : REAL;                   // 由卷径与圈数反推的等效厚度 [mm] / equivalent thickness reconstructed from diameter and revolutions [mm]
    uRollCount      : UDINT;                  // 累计换卷次数，饱和 [卷] / accumulated roll changes, saturating [roll]
    eErr            : UDINT;                  // 错误码，0=正常 / error id, 0=ok
    bError          : BOOL;                   // 故障标志，eErr 为故障级时 TRUE / error flag, TRUE on fault-level eErr
END_VAR
VAR
    fbTrigReset     : R_TRIG;                 // 复位上升沿实例，本体首部无条件刷新 / reset edge instance, refreshed unconditionally
    fbTrigNewRoll   : R_TRIG;                 // 换卷上升沿实例，本体首部无条件刷新 / new roll edge instance, refreshed unconditionally
    uLayerPrev      : UINT;                   // 上一拍层数，用于变化沿判定 [层] / previous layer count used by the edge test [layer]
    uLayerMaxEff    : UINT;                   // 钳位后的层数上限 [层] / clamped layer bound [layer]
    nLayerInt       : DINT;                   // 层数整数形态（截断）[层] / integer layer count, truncated [layer]
    fLayerFloat     : REAL;                   // 层数浮点形态 [层] / floating point layer count [layer]
    fRevAbs         : REAL;                   // 圈计数模长 [圈] / magnitude of the revolution count [rev]
    fDen            : REAL;                   // 等效厚度的反推分母（MAX(|圈|,1)）[圈] / denominator of the thickness estimate, at least one [rev]
    liRev           : LINT;                   // 圈计数升位副本（取模长前先升位）[圈] / widened revolution copy before taking the magnitude [rev]
    fDiaDelta       : REAL;                   // 卷径与芯径差 [mm] / diameter difference [mm]
    bInit           : BOOL := FALSE;          // 首扫标志，初值 FALSE，判据 NOT bInit / first-scan flag, initial FALSE, tested with NOT
END_VAR
VAR CONSTANT
    DL_WLC_LAYER_MIN : UINT := 10;            // 层数上限下限 [层] / layer bound lower limit [layer]
    DL_WLC_LAYER_MAX : UINT := 60000;         // 层数上限上限 [层] / layer bound upper limit [layer]
    DL_WLC_CNT_MAX   : UDINT := 16#FFFF_FFFE; // 换卷计数饱和值 [卷] / roll counter saturation value [roll]
    DL_WLC_TOL_LAYER : REAL := 1.0;           // 交叉校核容差 [层] / cross-check tolerance [layer]
    DL_WLC_ONE       : REAL := 1.0;           // 一值常量，分母下限与容差基底 [无量纲] / one constant used for the divisor floor [dimensionless]
    DL_WLC_TWO       : REAL := 2.0;           // 二值常量，层厚换算用 [无量纲] / two constant used by the thickness conversion [dimensionless]
    DL_FLOAT_EPS     : REAL := 1.0E-6;        // 浮点判等容差 [无量纲] / float equality tolerance [dimensionless]
    DL_WLC_INF_GUARD : REAL := 1.0E38;        // 非有限幅值判定阈值 [无量纲] / non-finite magnitude guard [dimensionless]
    DL_WLC_ZERO      : REAL := 0.0;           // 零值常量，避免裸字面量 [无量纲] / zero constant, avoids a bare literal [dimensionless]
    DL_WLC_CNT_ZERO  : UINT := 0;             // 无符号零常量 [无量纲] / unsigned zero constant [dimensionless]
    DL_WLC_LINT_ZERO : LINT := 0;             // LINT 零常量 [无量纲] / LINT zero constant [dimensionless]
END_VAR

// 段 1｜边沿实例无条件周期刷新（红线：严禁放入条件分支）/ segment 1, unconditional edge refresh
fbTrigReset(CLK := bReset);
fbTrigNewRoll(CLK := bNewRoll);

// 段 2｜输出与错误状态预置（层数与统计为保持量）/ segment 2, preset outputs, the counts are held
eErr := 0;                                    // 预置无错误 / preset no error
bError := FALSE;                              // 预置无故障 / preset no fault
bLayerEdge := FALSE;                          // 单周期脉冲先清 / clear the single-cycle pulse first
bInconsistent := FALSE;                       // 预置一致 / preset consistent

// 段 3｜首扫初始化（唯一合法范式：初值 FALSE，判据 NOT bInit）/ segment 3, first-scan initialisation
IF NOT bInit THEN
    uLayerDone := DL_WLC_CNT_ZERO;            // 首扫层数归 0 / layer count starts at zero
    uLayerPrev := DL_WLC_CNT_ZERO;            // 变化沿基准归 0 / the edge reference starts at zero
    uRollCount := 0;                          // 换卷统计清零 / clear the roll statistics
    fThicknessEst := DL_WLC_ZERO;             // 等效厚度清零 / clear the equivalent thickness
    bInit := TRUE;                            // 首扫只做一次 / first scan runs once only
END_IF

// 段 4｜复位沿：清零全部量（含累计统计）/ segment 4, reset clears everything
IF fbTrigReset.Q THEN
    uLayerDone := DL_WLC_CNT_ZERO;            // 层数清零 / clear the layer count
    uLayerPrev := DL_WLC_CNT_ZERO;            // 变化沿基准清零 / clear the edge reference
    uRollCount := 0;                          // 换卷统计清零 / clear the roll statistics
    fThicknessEst := DL_WLC_ZERO;             // 等效厚度清零 / clear the equivalent thickness
END_IF

// 段 5｜换卷沿：保留累计统计，只重置层数基准 / segment 5, a new roll keeps the statistics
IF fbTrigNewRoll.Q THEN
    uLayerDone := DL_WLC_CNT_ZERO;            // 新卷层数从 0 起 / a new roll starts at zero layers
    uLayerPrev := DL_WLC_CNT_ZERO;            // 变化沿基准重置 / reset the edge reference
    IF uRollCount < DL_WLC_CNT_MAX THEN
        uRollCount := uRollCount + 1;         // 饱和累计换卷次数 / saturating roll counter
    END_IF
END_IF

// 段 6｜使能闸：失能冻结层数 / segment 6, enable gate freezes the counts
IF NOT bEnable THEN
    RETURN;                                   // 失能即出口，输出保持 / disabled is the exit, the outputs are held
END_IF

// 段 7｜厚度与芯径闸（厚度在分母上，是除零唯一出口）/ segment 7, thickness and core gate
IF (fThickness <> fThickness) OR (fThickness <= DL_FLOAT_EPS) OR (fThickness > DL_WLC_INF_GUARD)
   OR (fCoreDiameter <> fCoreDiameter) OR (fCoreDiameter <= DL_FLOAT_EPS) THEN
    eErr := 16#0004_02E7;                     // 厚度或芯径非法故障码 / thickness or core fault id
    bError := TRUE;                           // 置故障标志 / raise the error flag
    RETURN;                                   // 故障级提前返回，层数冻结 / early return, the layer count is frozen
END_IF

// 段 8｜卷径闸（非有限或小于芯径，物理上不可能）/ segment 8, coil diameter gate
IF (fCoilDiameter <> fCoilDiameter) OR (fCoilDiameter > DL_WLC_INF_GUARD) OR (fCoilDiameter < fCoreDiameter) THEN
    eErr := 16#0004_02E8;                     // 卷径非法故障码 / illegal coil diameter fault id
    bError := TRUE;                           // 置故障标志 / raise the error flag
    RETURN;                                   // 故障级提前返回，层数冻结 / early return, the layer count is frozen
END_IF

// 段 9｜层数上限钳位（钳位后功能仍可用）/ segment 9, layer bound clamp
uLayerMaxEff := uLayerMax;                    // 取入参副本 / copy the input
IF uLayerMaxEff < DL_WLC_LAYER_MIN THEN
    uLayerMaxEff := DL_WLC_LAYER_MIN;         // 下限钳位 / clamp at the lower limit
    eErr := 16#0004_01D3;                     // 信息级：上限超域已钳位 / info level, the bound was clamped
ELSIF uLayerMaxEff > DL_WLC_LAYER_MAX THEN
    uLayerMaxEff := DL_WLC_LAYER_MAX;         // 上限钳位 / clamp at the upper limit
    eErr := 16#0004_01D3;                     // 信息级：上限超域已钳位 / info level, the bound was clamped
END_IF

// 段 10｜层数推算（分母已由段 7 保证 > 0）/ segment 10, layer computation
fDiaDelta := fCoilDiameter - fCoreDiameter;   // 卷径与芯径差 [mm] / diameter difference [mm]
fLayerFloat := fDiaDelta / (DL_WLC_TWO * fThickness); // 层数 = 差 / (2·厚度) [层] / layers equal the difference divided by twice the thickness [layer]
IF fLayerFloat > UINT_TO_REAL(uLayerMaxEff) THEN
    fLayerFloat := UINT_TO_REAL(uLayerMaxEff); // 超上限钳位 / clamp at the bound
    eErr := 16#0004_01D3;                     // 信息级：层数超上限已钳位 / info level, the layer count was clamped
END_IF
IF fLayerFloat < DL_WLC_ZERO THEN
    fLayerFloat := DL_WLC_ZERO;               // 卷径等于芯径时层数为 0 / a diameter equal to the core gives zero layers
END_IF
nLayerInt := REAL_TO_DINT(fLayerFloat);       // 截断取整为层数 [层] / truncate to an integer layer count [layer]
IF nLayerInt < 0 THEN
    nLayerInt := 0;                           // 防御性下界 / defensive floor
END_IF
uLayerDone := DINT_TO_UINT(nLayerInt);        // 发布已绕层数 [层] / publish the wound layer count [layer]

// 段 11｜剩余层数（下溢钳 0，绝不回绕）/ segment 11, remaining layers without underflow
IF uLayerDone >= uLayerMaxEff THEN
    uLayerRemain := DL_WLC_CNT_ZERO;          // 已到上限即剩余 0 / nothing remains at the bound
ELSE
    uLayerRemain := uLayerMaxEff - uLayerDone; // 剩余层数 [层] / remaining layers [layer]
END_IF

// 段 12｜交叉校核：圈计数取模长（先升 LINT 再取负，规避 DINT 最小值回绕）/ segment 12, cross-check
liRev := DINT_TO_LINT(diRevCount);            // 先升位，再取模长 / widen first, then take the magnitude
IF liRev < DL_WLC_LINT_ZERO THEN
    liRev := -liRev;                          // LINT 域取负安全 / negating inside LINT is safe
END_IF
fRevAbs := LINT_TO_REAL(liRev);               // 圈计数模长 [圈] / revolution magnitude [rev]
IF ABS(fLayerFloat - fRevAbs) > DL_WLC_TOL_LAYER THEN
    bInconsistent := TRUE;                    // 超过 1 层即提示（打滑/叠绕/噪声均可能）/ more than one layer apart is reported
    eErr := 16#0004_01D3;                     // 信息级：仅提示，不报故障（报故障会误停整线）/ info level only, a fault would stop the whole line
END_IF

// 段 13｜等效厚度反推（分母用 MAX(|圈|,1)，不用除零闸）/ segment 13, equivalent thickness
fDen := MAX(fRevAbs, DL_WLC_ONE);             // 圈数为 0 是开机常态，分母取下限 1 / zero revolutions is normal at start-up, use a floor of one
fThicknessEst := fDiaDelta / (DL_WLC_TWO * fDen); // 等效厚度 [mm] / equivalent thickness [mm]

// 段 14｜层数变化沿（单周期脉冲）/ segment 14, layer change edge
IF uLayerDone <> uLayerPrev THEN
    bLayerEdge := TRUE;                       // 层数变化即置单拍脉冲 / raise the single-cycle pulse on any change
    uLayerPrev := uLayerDone;                 // 更新比较基准 / update the reference
END_IF
END_FUNCTION_BLOCK
